(* IEC 61131-3 sources: daoli-st-library/DL_Process (part 25) *)

(* ---- FB_DL_CathodeKilnZoneSeq.st ---- *)
(*
  Component : FB_DL_CathodeKilnZoneSeq
  Category  : DL_Process
  Function  : 辊道窑多温区升温曲线执行状态机：预热→升温→保温→冷却→出料
  Complexity: C4
  开源溯源 : DLF 内部原创（R94 族模板派生）；参考语义来源见 SOURCE_HUNTING_MATRIX.md
  规则遵从 : R1-R16
  契约     : 输入 xStart 启动（上升沿启动，下降沿兼故障复位沿）、xStop 停止、xRollerOk 辊道运行正常、
             xRodBroken 断棒检测、xDischDone 出料完成、afZoneTempC 八温区实测温度定长数组 [℃]
             （ARRAY[0..7]，未用槽填零，R15 显式定长）、nZoneCount 有效温区数 [区]、
             rStartC 起始炉温 [℃]、rPreheatC 预热终点 [℃]、rSoakSetC 保温设定 [℃]、
             rRampRateKmin 升降温速率上限 [K/min]、rTempTolK 区温偏差允许带 [K]、
             rOverTempK 超温判据余量 [K]、rCoolTargetC 冷却终点 [℃]、rSoakTimeS 保温时间 [s]、
             rHeatMaxS 升温允许最长 [s]、rCoolMaxS 冷却允许最长 [s]、rDischTmoS 出料超时 [s]。
  输出     : 三路独立命令、ePhase 当前相、xFault/nFaultCode 故障、nWarnCode 信息级码、
             rZoneDevMaxK 各区相对保温设定的最大偏差 [K]、rMaxTempC/rMinTempC 区温极值 [℃]、
             xOverTemp 超温标志、xRateViol 速率越限标志。
  时序     : 同拍双窗配比约束 rHeatMaxS ≥ (rSoakSetC − rStartC) / rRampRateKmin × 60（否则升温窗
             先于工艺升温完成即超时）、rCoolMaxS ≥ (rSoakSetC − rCoolTargetC) / rRampRateKmin × 60。
  速率限幅 : 升温相以进相时刻的炉温为基准，允许温度 = 基准 + 速率 × 已用时间，实测超越即本拍断加热；
             降温相以进相时刻的炉温为基准，允许温度 = 基准 − 速率 × 已用时间，实测低于即本拍断风机。
  安全侧   : 断棒（xRodBroken）与辊道停转（NOT xRollerOk）在非待机相立即迁 FAULT 并撤销全部命令；
             断棒/停转在待机相不锁存，但阻断启动（启动条件已含两者）。
  复位沿   : 故障码锁存至 xStart 下降沿；复位后停在 IDLE，需重新给出启动上升沿才继续（不做自动再入）。
  码位     : 9820 升温速率超限（信息级）；9821 降温速率超限（信息级）；9822 区温偏差超带（信息级）；
             9823 超温转冷却（信息级）；9824 断棒（故障级）；9825 辊道停转（故障级）；
             9826 参数或温度数组非法（故障级）；9827 升温超时（故障级）；9828 冷却超时（故障级）；
             9829 出料超时（故障级）。信息级码一律不置 xFault。
*)
TYPE E_DL_KilnPhase :
(
    IDLE      := 0,    // 待机，全部命令撤销 EN: idle, every command withdrawn
    PREHEAT   := 10,   // 预热段升温 EN: the preheat ramp phase
    RAMP      := 20,   // 升温段至保温设定 EN: the ramp phase towards the soak setpoint
    SOAK      := 30,   // 保温段 EN: the soak phase
    COOL      := 40,   // 冷却段 EN: the cooling phase
    DISCHARGE := 50,   // 出料段 EN: the discharge phase
    FAULT     := 90    // 故障相，全部命令强制撤销 EN: fault phase, every command forced off
);
END_TYPE

FUNCTION_BLOCK FB_DL_CathodeKilnZoneSeq
VAR_INPUT
    xStart       : BOOL;                        // 启动（上升沿启动，下降沿复位故障） EN: start on the rising edge, reset the fault on the falling edge
    xStop        : BOOL;                        // 停止（任意相生效） EN: stop, effective in every phase
    xRollerOk    : BOOL;                        // 辊道运行正常（变频器运行反馈） EN: the roller table runs normally
    xRodBroken   : BOOL;                        // 断棒检测（安全侧信号） EN: the broken rod detection, a safety side signal
    xDischDone   : BOOL;                        // 出料完成（下游确认） EN: the discharge is complete, confirmed downstream
    afZoneTempC  : ARRAY[0..7] OF REAL;         // 八温区实测温度，未用槽填零 [℃] EN: the measured temperatures of eight zones, unused slots hold zero
    nZoneCount   : INT := 8;                    // 有效温区数 [区] EN: the number of valid zones
    rStartC      : REAL := 25.0;                // 起始炉温（升温速率基准的缺省值） [℃] EN: the starting furnace temperature used as the default ramp base
    rPreheatC    : REAL := 400.0;               // 预热终点温度 [℃] EN: the preheat end temperature
    rSoakSetC    : REAL := 800.0;               // 保温设定温度 [℃] EN: the soak setpoint temperature
    rRampRateKmin: REAL := 3.0;                 // 升降温速率上限 [K/min] EN: the upper bound of the heating and cooling rate
    rTempTolK    : REAL := 15.0;                // 区温偏差允许带 [K] EN: the allowed zone temperature deviation band
    rOverTempK   : REAL := 20.0;                // 超温判据余量（超过设定即转冷却） [K] EN: the over temperature margin above the setpoint
    rCoolTargetC : REAL := 80.0;                // 冷却终点温度 [℃] EN: the cooling end temperature
    rSoakTimeS   : REAL := 3600.0;              // 保温时间设定 [s] EN: the soak time setting
    rHeatMaxS    : REAL := 7200.0;              // 升温允许最长（预热+升温合计） [s] EN: the longest heating time covering preheat and ramp
    rCoolMaxS    : REAL := 7200.0;              // 冷却允许最长 [s] EN: the longest cooling time
    rDischTmoS   : REAL := 1800.0;              // 出料超时设定 [s] EN: the discharge timeout setting
END_VAR
VAR_OUTPUT
    xHeatCmd    : BOOL;               // 加热使能命令 EN: the heating enable command
    xFanCoolCmd : BOOL;               // 冷却风机命令 EN: the cooling fan command
    xDischCmd   : BOOL;               // 出料辊道命令 EN: the discharge conveyor command
    ePhase      : E_DL_KilnPhase;     // 当前相 EN: the current phase
    xFault      : BOOL;               // 故障标志（仅故障级码置位） EN: the fault flag, raised by fault class codes only
    nFaultCode  : INT;                // 故障码，锁存回放 EN: the fault code replayed from the latch
    nWarnCode   : INT;                // 信息级码（每拍重算） EN: the information class code recomputed every cycle
    rZoneDevMaxK: REAL;               // 各区相对保温设定的最大偏差 [K] EN: the largest zone deviation from the soak setpoint
    rMaxTempC   : REAL;               // 区温最大值 [℃] EN: the highest zone temperature
    rMinTempC   : REAL;               // 区温最小值 [℃] EN: the lowest zone temperature
    xOverTemp   : BOOL;               // 超温标志 EN: the over temperature flag
    xRateViol   : BOOL;               // 速率越限标志 EN: the rate violation flag
END_VAR
VAR
    tonHeat    : TON;                 // 升温（预热+升温）总时长定时器 EN: the total heating timer
    tonSoak    : TON;                 // 保温定时器 EN: the soak timer
    tonCool    : TON;                 // 冷却时长定时器 EN: the cooling timer
    tonDisch   : TON;                 // 出料超时定时器 EN: the discharge timeout
    fbStartRise: R_TRIG;              // xStart 上升沿（唯一启动沿） EN: the rising edge of xStart, the only start edge
    fbStartFall: F_TRIG;              // xStart 下降沿（复位沿） EN: the falling edge of xStart, the reset edge
    xFinAll    : BOOL;                // 标量浮点入参有限 EN: the scalar floating inputs are finite
    xZoneFin   : BOOL;                // 全部有效温区读数有限 EN: every valid zone reading is finite
    xParamBad  : BOOL;                // 参数或数组非法 EN: a parameter or the array is illegal
    xZoneDevOk : BOOL;                // 区温偏差在允许带内 EN: the zone deviation is inside the band
    i          : INT;                 // 温区循环索引 [区] EN: the zone loop index
    nScan      : INT;                 // 实际扫描温区数 [区] EN: the effective zone scan count
    rMax       : REAL;                // 区温最大值累加器 [℃] EN: the zone maximum accumulator
    rMin       : REAL;                // 区温最小值累加器 [℃] EN: the zone minimum accumulator
    rDev       : REAL;                // 偏差累加器 [K] EN: the deviation accumulator
    rDevMax    : REAL;                // 最大偏差 [K] EN: the largest deviation
    rHeatBaseC : REAL;                // 升温相进相基准炉温 [℃] EN: the furnace temperature latched when heating starts
    rCoolBaseC : REAL;                // 冷却相进相基准炉温 [℃] EN: the furnace temperature latched when cooling starts
    rAllowC    : REAL;                // 本拍允许温度（速率限幅） [℃] EN: the temperature allowed in this cycle by the rate limit
    rElapsedS  : REAL;                // 相内已用时间 [s] EN: the elapsed time inside the phase
    nMsSoak    : UDINT := 3600000;    // 保温毫秒数（缺省防零 PT） EN: the soak milliseconds, the default avoids a zero preset
    nMsHeat    : UDINT := 7200000;    // 升温毫秒数 EN: the heating milliseconds
    nMsCool    : UDINT := 7200000;    // 冷却毫秒数 EN: the cooling milliseconds
    nMsDisch   : UDINT := 1800000;    // 出料毫秒数 EN: the discharge milliseconds
    nCodeLatch : INT;                 // 故障码锁存副本 EN: the latched copy of the fault code
END_VAR
VAR CONSTANT
    DL_CKZ_Z      : REAL := 0.0;      // 浮点零常量 EN: the floating point zero constant
    DL_CKZ_SECMIN : REAL := 60.0;     // 分钟换算秒系数 EN: the minute to second factor
    DL_CKZ_K1000  : REAL := 1000.0;   // 秒转毫秒系数 EN: the second to millisecond factor
    DL_CKZ_IDX_MAX: INT := 7;         // 温区数组上界索引 [区] EN: the zone array upper bound index
    DL_CKZ_CNT_MAX: INT := 8;         // 温区个数上限 [区] EN: the zone count upper bound
    DL_CKZ_W_RATE : INT := 9820;      // 升温速率超限（信息级） EN: the heating rate violation, information class
    DL_CKZ_W_COOL : INT := 9821;      // 降温速率超限（信息级） EN: the cooling rate violation, information class
    DL_CKZ_W_DEV  : INT := 9822;      // 区温偏差超带（信息级） EN: the zone deviation violation, information class
    DL_CKZ_W_OVER : INT := 9823;      // 超温转冷却（信息级） EN: the over temperature transfer, information class
    DL_CKZ_C_ROD  : INT := 9824;      // 断棒（故障级） EN: the broken rod
    DL_CKZ_C_ROLL : INT := 9825;      // 辊道停转（故障级） EN: the roller table stopped
    DL_CKZ_C_PARAM: INT := 9826;      // 参数或温度数组非法（故障级） EN: a parameter or the temperature array is illegal
    DL_CKZ_C_HEAT : INT := 9827;      // 升温超时（故障级） EN: the heating timed out
    DL_CKZ_C_COOL : INT := 9828;      // 冷却超时（故障级） EN: the cooling timed out
    DL_CKZ_C_DISCH: INT := 9829;      // 出料超时（故障级） EN: the discharge timed out
END_VAR

// 段1｜参数与采样门禁：标量浮点闸 + 温区数组逐个闸（先判后用，换算在闸后）
xFinAll := (rStartC = rStartC) AND ((rStartC - rStartC) = DL_CKZ_Z)
        AND (rPreheatC = rPreheatC) AND ((rPreheatC - rPreheatC) = DL_CKZ_Z)
        AND (rSoakSetC = rSoakSetC) AND ((rSoakSetC - rSoakSetC) = DL_CKZ_Z)
        AND (rRampRateKmin = rRampRateKmin) AND ((rRampRateKmin - rRampRateKmin) = DL_CKZ_Z)
        AND (rTempTolK = rTempTolK) AND ((rTempTolK - rTempTolK) = DL_CKZ_Z)
        AND (rOverTempK = rOverTempK) AND ((rOverTempK - rOverTempK) = DL_CKZ_Z)
        AND (rCoolTargetC = rCoolTargetC) AND ((rCoolTargetC - rCoolTargetC) = DL_CKZ_Z)
        AND (rSoakTimeS = rSoakTimeS) AND ((rSoakTimeS - rSoakTimeS) = DL_CKZ_Z)
        AND (rHeatMaxS = rHeatMaxS) AND ((rHeatMaxS - rHeatMaxS) = DL_CKZ_Z)
        AND (rCoolMaxS = rCoolMaxS) AND ((rCoolMaxS - rCoolMaxS) = DL_CKZ_Z)
        AND (rDischTmoS = rDischTmoS) AND ((rDischTmoS - rDischTmoS) = DL_CKZ_Z);                        // 十一个标量入参有限性 EN: the finiteness of all eleven scalar inputs
xParamBad := (NOT xFinAll) OR (nZoneCount < 1) OR (nZoneCount > DL_CKZ_CNT_MAX)
          OR (rRampRateKmin <= DL_CKZ_Z) OR (rSoakTimeS <= DL_CKZ_Z) OR (rHeatMaxS <= DL_CKZ_Z)
          OR (rCoolMaxS <= DL_CKZ_Z) OR (rDischTmoS <= DL_CKZ_Z) OR (rTempTolK <= DL_CKZ_Z)
          OR (rOverTempK < DL_CKZ_Z) OR (rSoakSetC <= rPreheatC) OR (rPreheatC <= rStartC)
          OR (rCoolTargetC >= rSoakSetC);                                                                 // 域闸与曲线单调性约束 EN: the domain gate and the profile monotonicity
nScan := nZoneCount;                                                                                      // 扫描个数 [区] EN: the scan count
rMax := DL_CKZ_Z;                                                                                         // 最大值初值 [℃] EN: the maximum accumulator initial value
rMin := DL_CKZ_Z;                                                                                         // 最小值初值 [℃] EN: the minimum accumulator initial value
rDevMax := DL_CKZ_Z;                                                                                      // 最大偏差初值 [K] EN: the largest deviation initial value
xZoneFin := TRUE;                                                                                         // 假定温区有限 EN: assume the zones are finite
IF (nScan >= 1) AND (nScan <= DL_CKZ_CNT_MAX) THEN                                                       // 个数合法才访问数组 EN: access the array only with a legal count
    FOR i := 0 TO nScan - 1 DO                                                                           // 定长数组循环（上界已证 ≤7） EN: the fixed array loop, the bound is proven at most seven
        IF (i >= 0) AND (i <= DL_CKZ_IDX_MAX) THEN                                                       // 逐元素双边界校验 EN: the per element bound check
            IF (afZoneTempC[i] = afZoneTempC[i]) AND ((afZoneTempC[i] - afZoneTempC[i]) = DL_CKZ_Z) THEN
                IF (i = 0) OR (afZoneTempC[i] > rMax) THEN                                               // 首元素或更大值 EN: the first element or a larger value
                    rMax := afZoneTempC[i];                                                              // 更新最大值 [℃] EN: update the maximum
                END_IF
                IF (i = 0) OR (afZoneTempC[i] < rMin) THEN                                               // 首元素或更小值 EN: the first element or a smaller value
                    rMin := afZoneTempC[i];                                                              // 更新最小值 [℃] EN: update the minimum
                END_IF
                rDev := ABS(afZoneTempC[i] - rSoakSetC);                                                 // 相对保温设定的偏差 [K] EN: the deviation from the soak setpoint
                IF rDev > rDevMax THEN                                                                   // 取更大偏差 EN: keep the larger deviation
                    rDevMax := rDev;                                                                     // 更新最大偏差 [K] EN: update the largest deviation
                END_IF
            ELSE
                xZoneFin := FALSE;                                                                       // 记非有限元素 EN: mark the non finite element
            END_IF
        END_IF
    END_FOR
ELSE
    xZoneFin := FALSE;                                                                                   // 个数非法等同读数不可用 EN: an illegal count makes the readings unusable
END_IF
xParamBad := xParamBad OR (NOT xZoneFin);                                                                // 读数不可用并入参数闸（单点写入） EN: merge the unusable readings into the parameter gate
IF (NOT xParamBad) THEN                                                                                  // 参数合法才做时间换算 EN: convert only when the parameters are legal
    nMsSoak := REAL_TO_UDINT(rSoakTimeS * DL_CKZ_K1000);                                                 // 保温毫秒数 EN: the soak milliseconds
    nMsHeat := REAL_TO_UDINT(rHeatMaxS * DL_CKZ_K1000);                                                  // 升温毫秒数 EN: the heating milliseconds
    nMsCool := REAL_TO_UDINT(rCoolMaxS * DL_CKZ_K1000);                                                  // 冷却毫秒数 EN: the cooling milliseconds
    nMsDisch := REAL_TO_UDINT(rDischTmoS * DL_CKZ_K1000);                                                // 出料毫秒数 EN: the discharge milliseconds
END_IF
xZoneDevOk := (NOT xParamBad) AND (rDevMax <= rTempTolK);                                                // 区温偏差带内判据 EN: the zone deviation band test

// 段2｜四只定时器 + 两只边沿实例无条件周期刷新（CASE 内不调用实例）
tonHeat(IN := (ePhase = E_DL_KilnPhase.PREHEAT) OR (ePhase = E_DL_KilnPhase.RAMP), PT := UDINT_TO_TIME(nMsHeat));  // 升温总时长 EN: the total heating time
tonSoak(IN := (ePhase = E_DL_KilnPhase.SOAK) AND xZoneDevOk, PT := UDINT_TO_TIME(nMsSoak));                          // 保温计时（偏差在带内才累计） EN: count the soak only inside the band
tonCool(IN := (ePhase = E_DL_KilnPhase.COOL), PT := UDINT_TO_TIME(nMsCool));                                         // 冷却时长 EN: the cooling time
tonDisch(IN := (ePhase = E_DL_KilnPhase.DISCHARGE), PT := UDINT_TO_TIME(nMsDisch));                                  // 出料时长 EN: the discharge time
fbStartRise(CLK := xStart);                                                                                          // 启动沿 EN: the start edge
fbStartFall(CLK := xStart);                                                                                          // 复位沿 EN: the reset edge

// 段3｜输出预置（唯一预置点，CASE 内只置位；信息级码每拍重算）
xHeatCmd := FALSE;                        // 加热预置关 EN: preset the heating off
xFanCoolCmd := FALSE;                     // 风机预置停 EN: preset the fan off
xDischCmd := FALSE;                       // 出料预置停 EN: preset the discharge off
xFault := FALSE;                          // 故障标志预置假 EN: preset the fault flag false
nFaultCode := 0;                          // 故障码预置零 EN: preset the fault code to zero
nWarnCode := 0;                           // 信息码预置零 EN: preset the warning code to zero
xOverTemp := FALSE;                       // 超温标志预置假 EN: preset the over temperature flag false
xRateViol := FALSE;                       // 速率越限标志预置假 EN: preset the rate violation flag false
rZoneDevMaxK := rDevMax;                  // 最大偏差出口 [K] EN: publish the largest deviation
rMaxTempC := rMax;                        // 区温最大值出口 [℃] EN: publish the highest zone temperature
rMinTempC := rMin;                        // 区温最小值出口 [℃] EN: publish the lowest zone temperature

// 段4｜全局安全闸：参数非法 / 断棒 / 辊道停转 → 锁故障；xStop 撤销命令回待机
IF xParamBad THEN
    nCodeLatch := DL_CKZ_C_PARAM;                                                                        // 参数非法锁存 EN: latch the parameter code
    xFault := TRUE;                                                                                      // 置故障标志 EN: raise the fault flag
    nFaultCode := DL_CKZ_C_PARAM;                                                                        // 故障码出口 EN: publish the fault code
    ePhase := E_DL_KilnPhase.FAULT;                                                                      // 迁故障相 EN: move to the fault phase
ELSIF xRodBroken AND (ePhase <> E_DL_KilnPhase.IDLE) THEN
    nCodeLatch := DL_CKZ_C_ROD;                                                                          // 断棒锁存 EN: latch the broken rod code
    xFault := TRUE;                                                                                      // 置故障标志 EN: raise the fault flag
    nFaultCode := DL_CKZ_C_ROD;                                                                          // 故障码出口 EN: publish the fault code
    ePhase := E_DL_KilnPhase.FAULT;                                                                      // 迁故障相 EN: move to the fault phase
ELSIF (NOT xRollerOk) AND (ePhase <> E_DL_KilnPhase.IDLE) THEN
    nCodeLatch := DL_CKZ_C_ROLL;                                                                         // 辊道停转锁存 EN: latch the roller stop code
    xFault := TRUE;                                                                                      // 置故障标志 EN: raise the fault flag
    nFaultCode := DL_CKZ_C_ROLL;                                                                         // 故障码出口 EN: publish the fault code
    ePhase := E_DL_KilnPhase.FAULT;                                                                      // 迁故障相 EN: move to the fault phase
ELSIF xStop AND (ePhase <> E_DL_KilnPhase.IDLE) THEN
    ePhase := E_DL_KilnPhase.IDLE;                                                                       // 撤销型停车回待机 EN: a withdrawing stop returns to idle
END_IF

// 段5｜主状态机（ENUM + CASE，ELSE 兜底非法值）
IF ePhase <> E_DL_KilnPhase.FAULT THEN
CASE ePhase OF
E_DL_KilnPhase.IDLE:
    // 拍 N：待机；启动需辊道正常、无断棒、无停车（入相即锁存速率限幅基准炉温）
    IF fbStartRise.Q AND xRollerOk AND (NOT xRodBroken) AND (NOT xStop) AND (NOT xParamBad) THEN
        rHeatBaseC := rMax;                                                                              // 锁存升温基准炉温 [℃] EN: latch the heating base temperature
        ePhase := E_DL_KilnPhase.PREHEAT;                                                                // 本拍行为：进预热相 EN: enter the preheat phase
    END_IF

E_DL_KilnPhase.PREHEAT:
    // 拍 N：预热升温，速率越限即本拍断加热（信息级 9820），升到预热终点转升温相
    rElapsedS := TIME_TO_REAL(tonHeat.ET) * 0.001;                                                       // 已用时间 [s] EN: the elapsed time
    rAllowC := rHeatBaseC + rRampRateKmin * (rElapsedS / DL_CKZ_SECMIN);                                 // 允许温度 [℃] EN: the temperature allowed by the rate limit
    IF rMax > (rAllowC + rTempTolK) THEN                                                                 // 速率越限判据 EN: the rate violation test
        xRateViol := TRUE;                                                                               // 置越限标志 EN: raise the rate flag
        nWarnCode := DL_CKZ_W_RATE;                                                                      // 信息级码，不置故障 EN: an information class code, no fault
    ELSE
        xHeatCmd := TRUE;                                                                                // 加热允许 EN: heating allowed
    END_IF
    IF rMax >= rPreheatC THEN                                                                            // 预热到位 EN: the preheat is complete
        ePhase := E_DL_KilnPhase.RAMP;                                                                   // 本拍行为：进升温相 EN: enter the ramp phase
    ELSIF tonHeat.Q THEN
        nCodeLatch := DL_CKZ_C_HEAT;                                                                     // 升温超时 EN: the heating timed out
        xFault := TRUE;                                                                                  // 置故障标志 EN: raise the fault flag
        nFaultCode := DL_CKZ_C_HEAT;                                                                     // 故障码出口 EN: publish the fault code
        ePhase := E_DL_KilnPhase.FAULT;                                                                  // 迁故障相 EN: move to the fault phase
    END_IF

E_DL_KilnPhase.RAMP:
    // 拍 N：升温至保温设定，含速率限幅与升温超时兜底
    rElapsedS := TIME_TO_REAL(tonHeat.ET) * 0.001;                                                       // 已用时间（含预热相） [s] EN: the elapsed time including the preheat phase
    rAllowC := rHeatBaseC + rRampRateKmin * (rElapsedS / DL_CKZ_SECMIN);                                 // 允许温度 [℃] EN: the allowed temperature
    IF rMax > (rAllowC + rTempTolK) THEN                                                                 // 速率越限判据 EN: the rate violation test
        xRateViol := TRUE;                                                                               // 置越限标志 EN: raise the rate flag
        nWarnCode := DL_CKZ_W_RATE;                                                                      // 信息级码 EN: the information class code
    ELSE
        xHeatCmd := TRUE;                                                                                // 加热允许 EN: heating allowed
    END_IF
    IF rMax >= (rSoakSetC - rTempTolK) THEN                                                              // 到达保温窗口下沿 EN: reached the lower edge of the soak window
        ePhase := E_DL_KilnPhase.SOAK;                                                                   // 本拍行为：进保温相 EN: enter the soak phase
    ELSIF tonHeat.Q THEN
        nCodeLatch := DL_CKZ_C_HEAT;                                                                     // 升温超时 EN: the heating timed out
        xFault := TRUE;                                                                                  // 置故障标志 EN: raise the fault flag
        nFaultCode := DL_CKZ_C_HEAT;                                                                     // 故障码出口 EN: publish the fault code
        ePhase := E_DL_KilnPhase.FAULT;                                                                  // 迁故障相 EN: move to the fault phase
    END_IF

E_DL_KilnPhase.SOAK:
    // 拍 N：保温；超温立即转冷却（信息级 9823），偏差超带只告警（9822）且不累计保温时间
    IF rMax > (rSoakSetC + rOverTempK) THEN                                                              // 超温判据 EN: the over temperature test
        xOverTemp := TRUE;                                                                               // 置超温标志 EN: raise the over temperature flag
        nWarnCode := DL_CKZ_W_OVER;                                                                      // 超温信息级码 EN: the over temperature information code
        rCoolBaseC := rMin;                                                                              // 锁存冷却基准炉温 [℃] EN: latch the cooling base temperature
        ePhase := E_DL_KilnPhase.COOL;                                                                   // 本拍行为：立即转冷却 EN: transfer to cooling immediately
    ELSIF NOT xZoneDevOk THEN
        nWarnCode := DL_CKZ_W_DEV;                                                                       // 偏差超带告警（信息级） EN: warn about the zone deviation
        xHeatCmd := TRUE;                                                                                // 保持加热以拉回设定 EN: keep heating to recover the setpoint
    ELSE
        xHeatCmd := TRUE;                                                                                // 保温加热 EN: soak heating
        IF tonSoak.Q THEN                                                                                // 保温时间到 EN: the soak time elapsed
            rCoolBaseC := rMin;                                                                          // 锁存冷却基准炉温 [℃] EN: latch the cooling base temperature
            ePhase := E_DL_KilnPhase.COOL;                                                               // 本拍行为：进冷却相 EN: enter the cooling phase
        END_IF
    END_IF

E_DL_KilnPhase.COOL:
    // 拍 N：冷却；降温过快本拍断风机（信息级 9821），降到终点转出料，冷却超时判 9828
    rElapsedS := TIME_TO_REAL(tonCool.ET) * 0.001;                                                       // 冷却已用时间 [s] EN: the cooling elapsed time
    rAllowC := rCoolBaseC - rRampRateKmin * (rElapsedS / DL_CKZ_SECMIN);                                 // 允许温度（速率下限） [℃] EN: the allowed temperature floor
    IF rMin < (rAllowC - rTempTolK) THEN                                                                 // 降温超速率判据 EN: the over fast cooling test
        xRateViol := TRUE;                                                                               // 置越限标志 EN: raise the rate flag
        nWarnCode := DL_CKZ_W_COOL;                                                                      // 信息级码 EN: the information class code
    ELSE
        xFanCoolCmd := TRUE;                                                                             // 风机允许 EN: the fan is allowed
    END_IF
    IF rMax <= rCoolTargetC THEN                                                                         // 冷却到位 EN: the cooling is complete
        ePhase := E_DL_KilnPhase.DISCHARGE;                                                              // 本拍行为：进出料相 EN: enter the discharge phase
    ELSIF tonCool.Q THEN
        nCodeLatch := DL_CKZ_C_COOL;                                                                     // 冷却超时 EN: the cooling timed out
        xFault := TRUE;                                                                                  // 置故障标志 EN: raise the fault flag
        nFaultCode := DL_CKZ_C_COOL;                                                                     // 故障码出口 EN: publish the fault code
        ePhase := E_DL_KilnPhase.FAULT;                                                                  // 迁故障相 EN: move to the fault phase
    END_IF

E_DL_KilnPhase.DISCHARGE:
    // 拍 N：出料；下游确认回待机，超时判 9829（迁入本相已带参数闸复检）
    IF xDischDone THEN                                                                                   // 出料完成 EN: the discharge is complete
        ePhase := E_DL_KilnPhase.IDLE;                                                                   // 本拍行为：回待机 EN: back to idle
    ELSIF tonDisch.Q THEN
        nCodeLatch := DL_CKZ_C_DISCH;                                                                    // 出料超时 EN: the discharge timed out
        xFault := TRUE;                                                                                  // 置故障标志 EN: raise the fault flag
        nFaultCode := DL_CKZ_C_DISCH;                                                                    // 故障码出口 EN: publish the fault code
        ePhase := E_DL_KilnPhase.FAULT;                                                                  // 迁故障相 EN: move to the fault phase
    END_IF

E_DL_KilnPhase.FAULT:
    // 故障相（本段被外层 IF 排除，保留分支以满足枚举穷举）
    xFault := TRUE;                                                                                      // 保持故障标志 EN: keep the fault flag
    nFaultCode := nCodeLatch;                                                                            // 锁存回放 EN: replay the latch

ELSE
    // 非法状态兜底：绝不停在未知相
    nCodeLatch := DL_CKZ_C_PARAM;                                                                        // 非法状态归参数码 EN: treat an illegal state as a parameter code
    xFault := TRUE;                                                                                      // 置故障标志 EN: raise the fault flag
    nFaultCode := DL_CKZ_C_PARAM;                                                                        // 故障码出口 EN: publish the fault code
    ePhase := E_DL_KilnPhase.FAULT;                                                                      // 迁故障相 EN: move to the fault phase
END_CASE
END_IF

// 段6｜相独立使能出口（IDLE/FAULT 不置任何命令，天然强制撤销；出料相另给辊道命令）
CASE ePhase OF
E_DL_KilnPhase.DISCHARGE:
    xDischCmd := TRUE;                                                                                   // 出料辊道命令 EN: the discharge conveyor command
ELSE
    xDischCmd := FALSE;                                                                                  // 其余相撤销出料命令 EN: withdraw the discharge command elsewhere
END_CASE

// 段7｜故障相锁存回放 + 复位沿（xStart 下降沿清除，复位后停 IDLE 需重新给启动上升沿）
IF ePhase = E_DL_KilnPhase.FAULT THEN
    xFault := TRUE;                                                                                      // 故障标志保持 EN: keep the fault flag
    nFaultCode := nCodeLatch;                                                                            // 锁存回放，不按当下输入重推断 EN: replay the latch instead of re inferring
    nWarnCode := 0;                                                                                      // 故障相不报信息级码 EN: no information class code in the fault phase
    xHeatCmd := FALSE;                                                                                   // 加热强制关 EN: force the heating off
    xFanCoolCmd := FALSE;                                                                                // 风机强制停（断棒时避免热冲击） EN: force the fan off to avoid a thermal shock
    xDischCmd := FALSE;                                                                                  // 出料强制停 EN: force the discharge off
    IF fbStartFall.Q THEN
        nCodeLatch := 0;                                                                                 // 清除边：xStart 下降沿（头注释已声明） EN: clear on the falling edge of xStart
        ePhase := E_DL_KilnPhase.IDLE;                                                                   // 回待机 EN: back to idle
    END_IF
END_IF
END_FUNCTION_BLOCK

(* ---- FB_DL_CellAgingRestSeq.st ---- *)
(*
  组件名 Component   : FB_DL_CellAgingRestSeq
  子库 Sublibrary    : DL_Process
  版本 Version       : 1.0.0
  兼容性 Platform    : CODESYS 3.5 / TwinCAT 3 / 汇川 InoProShop / Machine Expert（仅 Standard.library）
  功能 Function      : 电芯老化静置顺控（自研行业池：锂电）：
                       1) 静置计时：tRestDur 总静置时长承载（独立 TON）；
                       2) 抽测窗口：静置相内周期开抽测窗（周期计 tonSampleInt 自复触，
                       R188），窗长 tSampleWin；窗口结束后锁存最后一次抽测值；
                       3) 时限到期判级出柜：静置时长到 → 按末次抽测电压与内阻判级
                       （合格 ePass / 降级 eMarginal / 不合格 eFail），结果锁存至复位；
                       4) 静置中断判据：抽测窗内电压越域持续 tVoltDevTo → 故障锁存。
  边界 Boundary      : ① 本件只出抽测请求与判级结论，不驱动充放电（老化柜本体自控）；
                       ② 判级只认末次抽测锁存值（禁按当下输入重推断，R152）；
                       ③ 周期窗计时自复触范式（R188），静置/窗口/越带确认独立实例；
                       ④ 故障锁存解除唯一路径 = bReset 上升沿（输入引脚，恒可达）；
                       ⑤ 无全局变量引用、无外部变量声明、无物理地址寻址。
  依赖 Depends       : Standard.library（R_TRIG / TON）
  溯源 Origin        : 道莅自研 clean-room（自研行业池：锂电老化静置共性语义，
                       零外部代码行复制）
  码位 Code          : 16#06_0_C0（Process 段 0006，C 子带 C0 格）
  码表 Error codes（本件格 06_0_C0，单轨子道：故障 0x02C0 / 信息 0x01C0）:
    16#0006_02C0 故障级：静置顺控故障总码（电压越域 / 组态非法 / 输入非有限），
                 锁存至复位
    16#0006_01C0 信息级：判级完成沿（ePass/eMarginal/eFail 写定拍）
  修订历史 Revision  :
    2026-11-19  v1.0.0  R44 首版（批次 4 · 序号 17）
*)

TYPE E_DL_CarPhase :
(
    eIdle     := 0,   // 空闲：未使能 / Idle, not enabled
    eRest     := 10,  // 静置：计时 + 周期抽测 / Resting with periodic sampling
    eSample   := 20,  // 抽测：窗口驻留 / Sampling window dwell
    eGrade    := 30,  // 判级：末次抽测定级 / Grading from last sample
    eDone     := 40,  // 完成：结论驻留 / Done, verdict held
    eFault    := 90   // 故障：总码锁存 / Fault, latched
);
END_TYPE

TYPE E_DL_CarGrade :
(
    eNone     := 0,   // 无结论 / No verdict
    ePass     := 10,  // 合格：电压内阻双达标 / Pass
    eMarginal := 20,  // 降级：电压入降级带 / Marginal
    eFail     := 30   // 不合格：越降级带下限或内阻不足 / Fail
);
END_TYPE

FUNCTION_BLOCK FB_DL_CellAgingRestSeq
VAR_INPUT
    bEnable     : BOOL;                  // 使能（电平）[-] / Enable
    bReset      : BOOL;                  // 上升沿清故障锁存 [-] / Reset edge
    fCellVoltV  : REAL;                  // 电芯实测电压 [伏特] / Cell voltage
    fIrMohm     : REAL;                  // 电芯实测内阻 [毫欧] / Internal resistance
    tRestDur    : TIME := T#72H;         // 总静置时长 [毫秒] / Total rest duration
    tSampleInt  : TIME := T#4H;          // 抽测周期 [毫秒] / Sample interval
    tSampleWin  : TIME := T#60S;         // 抽测窗口长 [毫秒] / Sample window duration
    fVoltPassLoV: REAL := 3.60;          // 合格电压下限 [伏特] / Pass voltage floor
    fVoltMargLoV: REAL := 3.50;          // 降级电压下限 [伏特] / Marginal voltage floor
    fIrMinMohm  : REAL := 1.0;           // 合格内阻下限 [毫欧] / IR pass floor
    tVoltDevTo  : TIME := T#10S;         // 电压越域确认窗 [毫秒] / Voltage deviation timeout
END_VAR
VAR_OUTPUT
    bSampleReq  : BOOL;                  // 抽测请求电平（窗口相）[-] / Sample request level
    fVoltLastV  : REAL;                  // 末次抽测电压 [伏特] / Last sampled voltage
    fIrLastMohm : REAL;                  // 末次抽测内阻 [毫欧] / Last sampled IR
    eGrade      : E_DL_CarGrade;         // 判级结论出口 / Grade verdict outlet
    ePhase      : E_DL_CarPhase;         // 相位出口，段尾单点映射 / Phase outlet
    bError      : BOOL;                  // 故障锁存标志 [-] / Fault latch flag
    uErrId      : UDINT;                 // 事件码，0 = 无事件 / Event code
END_VAR
VAR
    rtReset    : R_TRIG;                 // 复位沿实例，段 0 无条件刷新 / Reset edge
    tonRestDur : TON;                    // 静置总时长计时（独立实例） / Rest duration timer
    tonSampleInt: TON;                   // 抽测周期计（自复触，R188） / Sample interval timer
    tonSampleWin: TON;                   // 抽测窗口计时（独立实例） / Sample window timer
    tonVoltDevTo: TON;                   // 电压越域确认（专用超时件命名） / Voltage timeout
    _ePhase    : E_DL_CarPhase := E_DL_CarPhase.eIdle;    // 内部相位（CASE 唯一写入目标）/ Internal phase
    _eGrade    : E_DL_CarGrade := E_DL_CarGrade.eNone;    // 内部判级（锁存量）/ Internal grade
    _bFault    : BOOL;                   // 故障锁存位（锁存量） / Latched fault bit
    _uFault    : UDINT;                  // 故障码锁存（锁存量） / Latched fault code
    _bCfgBad   : BOOL;                   // 组态非法当拍量 [-] / Config illegal flag
    _bNonFin   : BOOL;                   // 输入非有限当拍量 [-] / Non-finite input flag
END_VAR
VAR CONSTANT
    DL_ABS_MAX : REAL := 1.0E30;         // 有限值判定上界 [工程单位] / Finite bound
    DL_ZERO    : REAL := 0.0;            // 零常量 [工程单位] / Zero constant
END_VAR

(* —— 段 0｜沿与定时器每拍无条件刷新（禁置于 IF/CASE 内；各实例独立禁复用） —— *)
rtReset(CLK := bReset);
tonRestDur (IN := (_ePhase = E_DL_CarPhase.eRest) AND (NOT _bFault), PT := tRestDur);
tonSampleInt(IN := (_ePhase = E_DL_CarPhase.eRest) AND (NOT _bFault) AND (NOT tonSampleInt.Q),
             PT := tSampleInt);          // 自复触周期窗：Q 拍断开一拍（R188）
tonSampleWin(IN := (_ePhase = E_DL_CarPhase.eSample) AND (NOT _bFault), PT := tSampleWin);
tonVoltDevTo(IN := (_ePhase = E_DL_CarPhase.eSample) AND ((fCellVoltV > fVoltPassLoV)
              OR (fCellVoltV < fVoltMargLoV)) AND (NOT _bFault), PT := tVoltDevTo);

(* —— 段 1｜瞬时量预清零（锁存量 _bFault/_uFault/_eGrade/fVoltLastV/fIrLastMohm 不入清单） —— *)
uErrId   := 16#0000_0000;
bSampleReq := FALSE;
_bCfgBad := FALSE;
_bNonFin := FALSE;

(* —— 段 2｜复位沿：故障与判级一次性清干净，相位回空闲 —— *)
IF rtReset.Q THEN
    _bFault := FALSE;
    _uFault := 16#0000_0000;
    _eGrade := E_DL_CarGrade.eNone;
    _ePhase := E_DL_CarPhase.eIdle;
END_IF

(* —— 段 3｜组态闸与非有限判据（覆盖全部参与判据换算引脚） —— *)
IF (fVoltMargLoV >= fVoltPassLoV) OR (fIrMinMohm <= DL_ZERO) OR (tRestDur = T#0S)
   OR (tSampleInt = T#0S) OR (tSampleWin = T#0S) OR (tVoltDevTo = T#0S) THEN
    _bCfgBad := TRUE;
END_IF
IF (fCellVoltV <> fCellVoltV) OR ((fCellVoltV - fCellVoltV) <> DL_ZERO)
   OR (fIrMohm <> fIrMohm) OR ((fIrMohm - fIrMohm) <> DL_ZERO) THEN
    _bNonFin := TRUE;
END_IF

(* —— 段 4｜主状态机：六态全覆盖 + ELSE 兜底 —— *)
CASE _ePhase OF

E_DL_CarPhase.eIdle:
    IF bEnable AND (NOT _bCfgBad) THEN
        _ePhase := E_DL_CarPhase.eRest;
    ELSIF bEnable AND _bCfgBad THEN
        _bFault := TRUE;
        _uFault := 16#0006_02C0;
        bError  := TRUE;
        _ePhase := E_DL_CarPhase.eFault;
    END_IF

E_DL_CarPhase.eRest:
    IF _bNonFin THEN
        _bFault := TRUE;
        _uFault := 16#0006_02C0;
        bError  := TRUE;
        _ePhase := E_DL_CarPhase.eFault;
    ELSIF NOT bEnable THEN
        _ePhase := E_DL_CarPhase.eIdle;  // 使能撤销回空闲
    ELSIF tonSampleInt.Q THEN
        _ePhase := E_DL_CarPhase.eSample;    // 抽测周期到：开抽测窗
    ELSIF tonRestDur.Q THEN
        _ePhase := E_DL_CarPhase.eGrade;     // 静置时长到：进判级相
    END_IF

E_DL_CarPhase.eSample:
    bSampleReq := TRUE;                  // 抽测请求电平（窗口相电平）
    IF _bNonFin THEN
        _bFault := TRUE;
        _uFault := 16#0006_02C0;
        bError  := TRUE;
        _ePhase := E_DL_CarPhase.eFault;
    ELSIF tonVoltDevTo.Q THEN
        _bFault := TRUE;                 // 窗内电压越域持续：锁存
        _uFault := 16#0006_02C0;
        bError  := TRUE;
        _ePhase := E_DL_CarPhase.eFault;
    ELSIF tonSampleWin.Q THEN
        fVoltLastV := fCellVoltV;        // 窗口结束：末次抽测值锁存（R152）
        fIrLastMohm := fIrMohm;
        bSampleReq := FALSE;
        _ePhase := E_DL_CarPhase.eRest;  // 回静置相（抽测周期重新起算）
    END_IF

E_DL_CarPhase.eGrade:
    (* 判级只认末次抽测锁存值（禁按当下输入重推断） *)
    IF (fVoltLastV >= fVoltPassLoV) AND (fIrLastMohm >= fIrMinMohm) THEN
        _eGrade := E_DL_CarGrade.ePass;  // 合格：双达标
    ELSIF (fVoltLastV >= fVoltMargLoV) AND (fIrLastMohm >= fIrMinMohm) THEN
        _eGrade := E_DL_CarGrade.eMarginal;      // 降级：电压入降级带
    ELSE
        _eGrade := E_DL_CarGrade.eFail;  // 不合格：越降级带或内阻不足
    END_IF
    uErrId := 16#0006_01C0;              // 信息级：判级完成沿
    _ePhase := E_DL_CarPhase.eDone;

E_DL_CarPhase.eDone:
    ;                                    // 结论锁存驻留（eGrade 出口回放），等复位或使能撤销
    IF NOT bEnable THEN
        _ePhase := E_DL_CarPhase.eIdle;  // 使能撤销回空闲（待机可返回路径）
    END_IF

E_DL_CarPhase.eFault:
    bError := TRUE;                      // 故障相驻留：判级与抽测值冻结，只认复位沿（段 2 迁出）
    ;                                    // （冻结语义：fVoltLastV/fIrLastMohm/_eGrade 保持）

ELSE
    _bFault := TRUE;                     // 兜底：非法相位锁存
    _uFault := 16#0006_02C0;
    bError  := TRUE;
    _ePhase := E_DL_CarPhase.eFault;
END_CASE

(* —— 段 5｜相位与判级出口单点映射（名实同源） —— *)
eGrade := _eGrade;
ePhase := _ePhase;
END_FUNCTION_BLOCK

(* ---- FB_DL_CellOcvBinSort.st ---- *)
(*
  FB_DL_CellOcvBinSort  —  OCV 分选档位落 bin（档位映射 + 满 bin 换道） / OCV bin sorting with grade mapping and full-bin lane change
  分类 Category : DL_Process
  版本 Version  : 1.0.0
  来源 Source   : roadmap-li-p1 — 锂电 OCV 分选工站真缺口
  溯源 Origin   : 道莅 clean-room 实现；四档电压阈值映射 + 落料计时 + 满 bin 换道停机为公开分选工艺逻辑，未复制任何源码行
  功能 Function : 1) 档位映射：fOcvMv 按 fTh1Mv~fTh4Mv 四阶梯阈值映射到档位 1~4
                  （阈值默认升序，第 4 档为 >= 阈值兜底档）；2) 落料相 eDispatch 由 tDrop 计时；
                  3) 档位 bin 计数 nBinUsed[档位] 递增，达 nBinCap 即 bBinFull 置位并在
                  段 3 以 03A1 锁存（满 bin 换道请求，须人工清空后复位）；
                  4) 故障级单码 03A1，归因由 eCause 独立成员承载（R190）；
                  5) 信息级 04C9 = 单件分选完成沿；6) 解除式全当拍量（R240）。
  接口 Interface: 输入 OCV 电压 + 四阈 + 容量 + 落料时间；输出状态/档位/各 bin 计数/码
  边界 Boundary : ① 组态闸：四阈值非严格升序（fTh2Mv <= fTh1Mv 等）、nBinCap = 0、
                  tDrop <= T#0S 任一成立 → 03A1 锁存；
                  ② 档位数组下标写前显式钳制（nGrade 落在 1..4，越界不写，ELSE 兜底归 4 档）；
                  ③ 浮点阈值判据为「>=」单侧直比（阈值本身无容差语义，避免误判），电压量纲
                  mV 整数化输入；④ 落料 TON 与 R_TRIG 段 0 无条件周期调用；
                  ⑤ 故障相迁出唯一路径 = bReset 上升沿；⑥ 零全局耦合（无 GVL / %I %Q %M）。
  依赖 Depends  : Standard.library（TON / R_TRIG）
  码表 Error codes（Process 段 0005，故障窗口 03A1 / 信息窗口 04C9）:
    16#0005_03A1 故障级：分选故障总码（组态非法 / 落料超时 / 目标 bin 已满需换道），
                 锁存至 bReset 上升沿；归因见 eCause，不新增码位（派单硬约束单码）
    16#0005_04C9 信息级：单件分选完成沿（落料完成计数后单拍）
  修订历史 Revision :
    2026-11-19  v1.0.0  R43 首版（批次 1 · 序号 5）
*)

TYPE E_DL_OcvState :
(
    eIdle     := 0,   // 未使能待启动 / Idle, waiting start
    eClassify := 10,  // 档位判定中 / Grade classification
    eDispatch := 20,  // 落料中（落料计时） / Dispatching with drop timer
    eDone     := 50,  // 单件完成 / Single piece done
    eFault    := 90   // 故障锁存相 / Fault latched phase
);
END_TYPE

TYPE E_DL_OcvCause :
(
    eNone       := 0, // 无故障成因 / No cause
    eCfgIllegal := 1, // 组态非法 / Illegal configuration
    eDropTmo    := 2, // 落料超时 / Drop timeout
    eBinFull    := 3  // 目标 bin 已满（换道请求） / Target bin full, lane change
);
END_TYPE

FUNCTION_BLOCK FB_DL_CellOcvBinSort
VAR_INPUT
    fOcvMv      : REAL := 0.0;        // 单体 OCV 电压 [mV] / Cell OCV voltage
    fTh1Mv      : REAL := 3300.0;     // 1/2 档分界阈值 [mV] / Grade 1-2 threshold
    fTh2Mv      : REAL := 3350.0;     // 2/3 档分界阈值 [mV] / Grade 2-3 threshold
    fTh3Mv      : REAL := 3400.0;     // 3/4 档分界阈值 [mV] / Grade 3-4 threshold
    fTh4Mv      : REAL := 3450.0;     // 4 档上界（>= 归 4 档） [mV] / Grade 4 upper threshold
    nBinCap     : UINT := 500;        // 单 bin 容量 [件]，域 > 0 / Bin capacity
    tDrop       : TIME := T#800MS;    // 落料时长 [ms]，域 > 0 / Drop duration
    bStart      : BOOL := FALSE;      // 启动命令（电平）[-] / Start command
    bBinCleared : BOOL := FALSE;      // bin 已清空确认（电平）[-] / Bin cleared acknowledge
    bReset      : BOOL := FALSE;      // 复位命令，上升沿清故障 [-] / Reset edge
END_VAR
VAR_OUTPUT
    eState      : E_DL_OcvState;      // 状态出口，段 6 单点映射 / State outlet
    eCause      : E_DL_OcvCause;      // 故障成因出口（R190） / Fault cause outlet
    nGrade      : UINT;               // 当前档位 0~4，0 = 未判定 / Current grade
    anBinUsed   : ARRAY[1..4] OF UDINT;   // 各档 bin 已用计数 [件] / Per-grade bin usage
    bBinFull    : BOOL;               // 满 bin 标志镜像 [-] / Bin full mirror
    bCycleDone  : BOOL;               // 单件完成标志 [-] / Piece done flag
    bError      : BOOL;               // 故障锁存标志 [-] / Fault latch flag
    nErrId      : UDINT;              // 事件码，0 = 无事件 / Event code
END_VAR
VAR
    _eState     : E_DL_OcvState := E_DL_OcvState.eIdle;   // 内部相位（CASE 唯一写入目标） / Internal phase
    _eCause     : E_DL_OcvCause := E_DL_OcvCause.eNone;   // 故障成因锁存（锁存量） / Latched cause
    tonDrop     : TON;                // 落料计时实例，每周期无条件调用 / Drop timer
    rtReset     : R_TRIG;             // 复位沿实例，每周期无条件调用 / Reset edge
    _anBinUsed  : ARRAY[1..4] OF UDINT;   // 内部 bin 计数（持久，段 6 映射） / Internal bin usage
    _nGrade     : UINT;               // 档位判定结果（当拍量） / Grade verdict
    _bCfgBad    : BOOL;               // 组态非法当拍量 [-] / Config illegal
    _bFault     : BOOL;               // 故障锁存位（锁存量） / Latched fault bit
    _uFault     : UDINT;              // 故障码锁存（锁存量） / Latched fault code
    _uInfo      : UDINT;              // 信息码，每拍重算 / Transient info code
END_VAR

(* —— 段 0：沿实例与定时器无条件周期刷新 + 档位判定（纯函数式，无副作用） —— *)
IF fOcvMv < fTh1Mv THEN                        // 低于 1/2 分界：1 档 / Below first threshold: grade 1
    _nGrade := 1;
ELSIF fOcvMv < fTh2Mv THEN                     // 低于 2/3 分界：2 档 / Grade 2
    _nGrade := 2;
ELSIF fOcvMv < fTh3Mv THEN                     // 低于 3/4 分界：3 档 / Grade 3
    _nGrade := 3;
ELSE                                           // 兜底：>= 3/4 分界归 4 档 / Fallback grade 4
    _nGrade := 4;
END_IF
_bCfgBad := (fTh2Mv <= fTh1Mv) OR (fTh3Mv <= fTh2Mv) OR (fTh4Mv <= fTh3Mv)
            OR (nBinCap = 0) OR (tDrop <= T#0S);                   // 组态非法当拍量 / Config illegal
rtReset(CLK := bReset);                                            // 复位沿，每拍必调 / Reset edge
tonDrop(IN := (_eState = E_DL_OcvState.eDispatch), PT := tDrop);   // 落料计时 / Drop timer

(* —— 段 1：单拍量预清零（锁存量与 bin 计数均不入清单） —— *)
_uInfo := 16#0000_0000;            // 信息码每拍重算 / Info recomputed
nGrade := 0;                       // 档位出口缺省 0 / Grade default
bBinFull := FALSE;                 // 满 bin 镜像缺省 FALSE / Bin full default
bCycleDone := FALSE;               // 完成标志缺省 FALSE / Done default
nErrId := 16#0000_0000;            // 事件码缺省无事件 / Event code default

(* —— 段 2：复位沿 + 组态域闸 —— *)
IF rtReset.Q THEN                              // rtReset.Q = 当拍量 / current scan
    _bFault := FALSE;                          // 清故障锁存位（锁存量） / Clear fault latch
    _uFault := 16#0000_0000;                   // 清故障锁存码（锁存量） / Clear fault code
    _eCause := E_DL_OcvCause.eNone;            // 清成因（锁存量） / Clear cause
    IF _eState = E_DL_OcvState.eFault THEN
        _eState := E_DL_OcvState.eIdle;        // 故障相迁出：回未使能 / Fault exit to idle
    END_IF
END_IF
IF _bCfgBad THEN                               // 组态域闸 / Config gate
    _uFault := 16#0005_03A1;                   // 故障级：分选故障总码 / Process fault code
    _eCause := E_DL_OcvCause.eCfgIllegal;      // 归因：组态非法 / Cause: illegal config
    _bFault := TRUE;                           // 标志与码位配对（R45） / Flag paired with code
END_IF

(* —— 段 3：落料超时与满 bin 换道（判据当拍量；下标写前钳制） —— *)
IF (NOT _bFault) AND tonDrop.Q THEN            // 落料超时 / Drop timeout
    _uFault := 16#0005_03A1;
    _eCause := E_DL_OcvCause.eDropTmo;         // 归因：落料超时 / Cause: drop timeout
    _bFault := TRUE;
END_IF
IF (NOT _bFault) AND (_nGrade >= 1) AND (_nGrade <= 4)
   AND (_anBinUsed[_nGrade] >= nBinCap) AND (NOT bBinCleared) THEN   // 目标 bin 已满且未清空 / Target bin full
    _uFault := 16#0005_03A1;
    _eCause := E_DL_OcvCause.eBinFull;         // 归因：满 bin 换道 / Cause: bin full
    _bFault := TRUE;
END_IF

(* —— 段 4：故障解除式（R240；全当拍量）：rtReset.Q / NOT _bCfgBad / NOT tonDrop.Q / bBinCleared —— *)
IF rtReset.Q AND (NOT _bCfgBad) AND (NOT tonDrop.Q) AND bBinCleared THEN
    _bFault := FALSE;                          // 清故障锁存位（锁存量） / Clear fault latch
    _uFault := 16#0000_0000;                   // 清故障锁存码（锁存量） / Clear fault code
    _eCause := E_DL_OcvCause.eNone;            // 清成因（锁存量） / Clear cause
END_IF

(* —— 段 4A：故障锁存相位迁移闸 —— *)
IF _bFault AND (_eState <> E_DL_OcvState.eFault) THEN
    _eState := E_DL_OcvState.eFault;           // 锁存即入故障相 / Latch enters fault phase
END_IF

(* —— 段 5：相位机（CASE 全覆盖 + ELSE 兜底） —— *)
CASE _eState OF

E_DL_OcvState.eIdle:
    IF bStart AND (NOT _bFault) THEN           // 启动条件 / Start gate
        _eState := E_DL_OcvState.eClassify;    // 进档位判定相 / Enter classification
    END_IF

E_DL_OcvState.eClassify:
    IF (_nGrade >= 1) AND (_nGrade <= 4) THEN  // 出口 1：档位有效（下标已钳制） / Valid grade
        _eState := E_DL_OcvState.eDispatch;    // 进落料相 / Enter dispatch
    ELSIF NOT bStart THEN                      // 出口 2：撤启动（R98 双出口） / Start released
        _eState := E_DL_OcvState.eIdle;
    END_IF

E_DL_OcvState.eDispatch:
    IF tonDrop.Q THEN                          // 落料到时 / Drop elapsed
        IF (_nGrade >= 1) AND (_nGrade <= 4) AND (NOT (_anBinUsed[_nGrade] >= nBinCap)) THEN
            _anBinUsed[_nGrade] := _anBinUsed[_nGrade] + 1;   // 计数递增（钳制下标 + 容量复核） / Increment with clamped index
        END_IF
        _uInfo := 16#0005_04C9;                // 信息级：单件分选完成沿 / Info: piece sorted edge
        _eState := E_DL_OcvState.eDone;        // 进完成相 / Enter done
    ELSIF NOT bStart THEN                      // 撤启动：中止 / Abort
        _eState := E_DL_OcvState.eIdle;
    END_IF

E_DL_OcvState.eDone:
    IF NOT bStart THEN                         // 撤启动回空闲 / Start released returns idle
        _eState := E_DL_OcvState.eIdle;
    END_IF

E_DL_OcvState.eFault:
    ;                                          // 故障相：仅段 4 复位沿可迁出 / Only reset exits

ELSE
    _uFault := 16#0005_03A1;                   // 故障级：非法相位兜底（归并总码） / Illegal phase fallback
    _eCause := E_DL_OcvCause.eCfgIllegal;      // 归因：相位非法归并组态 / Cause: phase illegal
    _bFault := TRUE;
    _eState := E_DL_OcvState.eFault;           // 强制回故障相 / Force fault phase

END_CASE

(* —— 段 6：出口单点映射（名实同源；锁存码回放） —— *)
nGrade := _nGrade;                             // 档位出口 / Grade outlet
anBinUsed[1] := _anBinUsed[1];                 // 1 档计数映射 / Grade 1 usage
anBinUsed[2] := _anBinUsed[2];                 // 2 档计数映射 / Grade 2 usage
anBinUsed[3] := _anBinUsed[3];                 // 3 档计数映射 / Grade 3 usage
anBinUsed[4] := _anBinUsed[4];                 // 4 档计数映射 / Grade 4 usage
bBinFull := (_nGrade >= 1) AND (_nGrade <= 4) AND (_anBinUsed[_nGrade] >= nBinCap);  // 满 bin 镜像 / Bin full mirror
bCycleDone := (_eState = E_DL_OcvState.eDone);// 完成标志 / Done flag
IF _bFault THEN
    nErrId := _uFault;                         // 故障锁存码回放 / Replay latched code
ELSE
    nErrId := _uInfo;                          // 信息码 / Transient info
END_IF
bError := _bFault;                             // 故障标志同源 / Flag from latch
eState := _eState;                             // 状态出口 / State outlet
eCause := _eCause;                             // 成因出口 / Cause outlet

END_FUNCTION_BLOCK

(* ---- FB_DL_CellSortingBin.st ---- *)
(*==============================================================================
 * 组件名称 (Component)  : FB_DL_CellSortingBin
 * 所属子库 (Sublibrary) : DL_Process
 * 当前版本 (Version)    : 1.0.0
 * 兼容性   (Platform)   : CODESYS 3.5+ / TwinCAT 3 / 汇川 InoProShop / 施耐德 Machine Expert
 *                         仅依赖 Standard.library（R_TRIG），零厂商私有库
 * 功能描述 (Function)   : 电池片分选落料 + 料仓满溢调度。
 *                           ① 档位→料仓映射：anGradeMap[nGrade − 1] 给出目标仓号，−1 表示该档
 *                              "不落料"（工艺上存在 NG 档直接走废料带、不进分选仓的情形）。
 *                           ② 满溢调度：目标仓已满（anBinCount ≥ anBinCapacity）时**不丢片**，
 *                              自动旁路到备仓 nBackupBin，并置 bOverflowBypass 锁存告警
 *                              （旁路是被动降级，必须让维护看见；悄悄丢片是最坏结果）。
 *                           ③ 双满兜底：目标仓与备仓同时满 → bNoBin 锁存故障、不落料、
 *                              由上层停机或切换收料框（本件不擅自选第三个仓——仓序属产线配置，
 *                              不是算法可以推断的）。
 *                           ④ 计数在**成功落料后**自增（inc-place 写回调用方的 anBinCount），
 *                              杜绝"先计数后落料"导致的仓位数虚高。
 * 接口     (Interface)  : 输入 nGrade 当前档位（1..8）、bDropCmd 落料命令（上升沿执行）、
 *                         anBinCount 各仓当前计数（VAR_IN_OUT，成功落料后自增）、
 *                         anBinCapacity 各仓容量（配置）、anGradeMap 档位到料仓映射（配置，−1 不落）、
 *                         nBackupBin 备仓号、bReset 复位；输出 nTargetBin 目标仓（−1 无）、
 *                         bDrop 落料脉冲（单拍）、bOverflowBypass 旁路告警（锁存）、
 *                         bNoBin 无可用仓（锁存）、bGradeUnmapped 该档不落料（当拍量）、
 *                         eState / eCause / bError。
 * 边界     (Boundary)   : ① **属主边界（写死）：本件只做"档位到仓号的选择与满溢旁路"，
 *                         不驱动气缸/翻转机构、不做到位确认**。执行机构动作与到位联锁属
 *                         落料执行 POU（可复用 `I_DL_Cylinder` 族）；本件只出目标仓号与落料脉冲。
 *                         ② 组态闸：nGrade < 1 或 > 8（越映射表边界）、nBackupBin 越 0..3、
 *                         任一 anBinCapacity[i] <= 0、映射表值 > 3（越仓边界）或 < −1、
 *                         映射表指向的仓不存在 → 故障锁存，落料脉冲不出（宁可不落，不可乱落）。
 *                         ③ 4 仓定长（ARRAY[0..3]）、8 档定长（ARRAY[0..7]）：容量写死在类型里，
 *                         改仓数须改类型定义，不允许"运行期可变长度"（那会越界）。
 *                         ④ 单枚 R_TRIG（bDropCmd）+ 单枚 R_TRIG（bReset）段 0 无条件周期刷新；
 *                         无 TON，故无跨相复位风险。
 *                         ⑤ 故障相与旁路锁存迁出唯一路径 = bReset 上升沿（R228B）。
 *                         ⑥ 零全局耦合（无 GVL / 无 VAR_EXTERNAL / 无物理地址）。
 * 分工声明 (Scope)      : 与 `FB_DL_Cylinder` 族（执行机构）分工——本件是**调度/记账**件，
 *                         输出仓号与脉冲；执行件负责把片真送进仓。二者不可混写在一个 FB 里，
 *                         否则换执行机构时要重测记账逻辑。
 * 来源标签 (Source Tag) : ROADMAP B 类（光伏电池片分选落料，自研 clean-room，无外源代码）
 * 解除式   (Release)    : bReset 上升沿 ∧ 组态合法 → 清 bNoBin / bOverflowBypass 锁存。
 *                         自证可满足：清仓（计数减少）或复位后即解除，无恒假因子。
 * 码表     (Codes)      : 本件不占用任何全局数字码位。出口为 INT 仓号 + BOOL 组 + ENUM
 *                         （eState / eCause）；数字码位待主控收口阶段统一派号。
 * 红线自检 (Redline)    : R1 ✓ 零 GVL/VAR_EXTERNAL ｜ R2 ✓ 零 %I/%Q/%M ｜ R3 ✓ 纯 IEC 61131-3
 *                         R4 ✓ 数组边界闸 + 映射值域闸 + 容量非正闸 ｜ R5 ✓ 声明逐行同行双语注释
 *                         R6 ✓ ENUM+CASE 含 ELSE ｜ R7 ✓ R_TRIG 段 0 无条件刷新
 * 修订历史 (Revision)   : 2026-11-19  v1.0.0  R46 首版（批次 3 · 序号 14）
 *==============================================================================*)

TYPE E_DL_CsbState :
(
    eIdle  := 0,    // 等待落料命令 / Awaiting a drop command
    eRun   := 10,   // 正常落料运行相 / Normal dropping
    eBypass:= 20,   // 满溢旁路相（走备仓，告警保持） / Overflow bypass phase
    eFault := 90    // 无可用仓/组态故障相 / No-bin or configuration fault
);
END_TYPE

TYPE E_DL_CsbCause :
(
    eNone        := 0,   // 无异常 / No anomaly
    eCfgIllegal  := 1,   // 组态非法（映射/容量/备仓越界） / Illegal configuration
    eOverflow    := 2,   // 目标仓满溢，已旁路到备仓 / Target bin full, bypassed to the backup bin
    eNoBin       := 3,   // 目标仓与备仓同时满，无可用仓 / Target and backup both full
    eGradeUnmapped:= 4,  // 该档不落料（映射为 −1） / Grade intentionally not dropped
    ePhaseBad    := 5    // 非法相位兜底 / Illegal phase fallback
);
END_TYPE

FUNCTION_BLOCK FB_DL_CellSortingBin
VAR_IN_OUT
    anBinCount : ARRAY[0..3] OF DINT;       // 各仓当前计数（成功落料后本件自增） [片] / Bin counts, incremented by this unit on success [pcs]
END_VAR
VAR_INPUT
    nGrade        : INT := 1;               // 当前档位，域 1..8 / Present grade, 1..8
    bDropCmd      : BOOL := FALSE;          // 落料命令，上升沿执行一次 [-] / Drop command, acts once per rising edge
    anBinCapacity : ARRAY[0..3] OF DINT;    // 各仓容量（配置），每项域 > 0 [片] / Bin capacities, each > 0 [pcs]
    anGradeMap    : ARRAY[0..7] OF INT;     // 档位到仓映射（配置），值域 −1 或 0..3 [-] / Grade-to-bin map, -1 or 0..3
    nBackupBin    : INT := 3;               // 备仓号，域 0..3 / Backup bin index, 0..3
    bReset        : BOOL := FALSE;          // 复位，上升沿清旁路与无仓锁存 [-] / Reset, rising edge clears latches
END_VAR
VAR_OUTPUT
    nTargetBin      : INT;                  // 本拍目标仓号，−1 表示无 / Target bin this scan, -1 means none
    bDrop           : BOOL;                 // 落料脉冲（单拍） [-] / Drop pulse, single scan
    bOverflowBypass : BOOL;                 // 满溢旁路告警（锁存） [-] / Overflow bypass alarm, latched
    bNoBin          : BOOL;                 // 无可用仓（锁存故障） [-] / No available bin, latched fault
    bGradeUnmapped  : BOOL;                 // 该档不落料（当拍量，非故障） [-] / Grade not dropped, per scan, not a fault
    eState          : E_DL_CsbState;        // 状态出口 [-] / State outlet
    eCause          : E_DL_CsbCause;        // 成因出口（R190 归因唯一） [-] / Cause outlet
    bError          : BOOL;                 // 故障标志（无仓/组态非法；旁路不算故障） [-] / Error flag, bypass is not a fault
END_VAR
VAR
    _eState   : E_DL_CsbState := E_DL_CsbState.eIdle;    // 内部相位（CASE 唯一写入目标） / Internal phase
    _eCause   : E_DL_CsbCause := E_DL_CsbCause.eNone;    // 成因锁存量 / Latched cause
    rtDrop    : R_TRIG;                 // 落料命令沿实例，段 0 无条件调用 / Drop edge instance
    rtReset   : R_TRIG;                 // 复位沿实例，段 0 无条件调用 / Reset edge instance
    _bBypass  : BOOL;                   // 旁路告警锁存位（锁存量） / Latched bypass alarm
    _bNoBin   : BOOL;                   // 无可用仓锁存位（锁存量） / Latched no-bin fault
    _bCfgBad  : BOOL;                   // 组态非法当拍量 [-] / Illegal configuration this scan
    _bMapBad  : BOOL;                   // 映射表非法当拍量 [-] / Illegal map this scan
    _nBin     : INT;                    // 映射得到的目标仓号中间量 [-] / Mapped target bin intermediate
    _nMapIdx  : INT;                    // 映射查表索引（已钳位） [-] / Clamped map index
    _i        : INT;                    // 遍历索引 / Loop index
END_VAR
VAR CONSTANT
    DL_CSB_BINMAX : INT := 3;           // 仓号上界（与 ARRAY[0..3] 一致） [仓] / Bin index bound matching the array
    DL_CSB_GRDMAX : INT := 8;           // 档位上界（与 ARRAY[0..7] 一致） [档] / Grade bound matching the array
    DL_CSB_NOBIN  : INT := -1;          // 无目标仓哨兵值 [-] / Sentinel for "no target bin"
END_VAR

(* —— 段 0：组态闸派生 + 两沿实例无条件周期刷新 —— *)
_bMapBad := FALSE;                                          // 映射非法初值 / Map-illegal initial value
FOR _i := 0 TO DL_CSB_GRDMAX - 1 DO
    IF (anGradeMap[_i] > DL_CSB_BINMAX) OR (anGradeMap[_i] < DL_CSB_NOBIN) THEN
        _bMapBad := TRUE;                                   // 映射值越界（> 3 或 < −1） / Map value out of range
    END_IF
END_FOR
FOR _i := 0 TO DL_CSB_BINMAX DO
    IF anBinCapacity[_i] <= 0 THEN
        _bMapBad := TRUE;                                   // 容量非正（永不装满或立即装满，皆病态） / Non-positive capacity is degenerate
    END_IF
END_FOR
_bCfgBad := _bMapBad
        OR (nBackupBin < 0) OR (nBackupBin > DL_CSB_BINMAX)   // 备仓号越界 / Backup index out of range
        OR (nGrade < 1) OR (nGrade > DL_CSB_GRDMAX);          // 档位越映射表边界 / Grade out of the map bounds
rtDrop(CLK := bDropCmd);                                    // 落料沿，每拍必调（R228A） / Drop edge, every scan
rtReset(CLK := bReset);                                     // 复位沿，每拍必调 / Reset edge, every scan

(* —— 段 1：单拍量预清零（锁存量 _bBypass / _bNoBin / _eCause 不入清单，R107） —— *)
nTargetBin     := DL_CSB_NOBIN;     // 目标仓缺省无 / Target bin defaults to none
bDrop          := FALSE;            // 落料脉冲每拍预清 / Drop pulse preset
bOverflowBypass:= FALSE;            // 旁路出口每拍预清 / Bypass outlet preset
bNoBin         := FALSE;            // 无仓出口每拍预清 / No-bin outlet preset
bGradeUnmapped := FALSE;            // 不落料标志每拍预清 / Unmapped flag preset
bError         := FALSE;            // 故障标志每拍预清（R45 配对） / Error flag preset

(* —— 段 2：复位沿 + 组态闸 —— *)
IF rtReset.Q THEN
    _bBypass := FALSE;                                  // 清旁路告警锁存 / Clear the bypass alarm
    _bNoBin  := FALSE;                                  // 清无仓锁存 / Clear the no-bin latch
    _eCause  := E_DL_CsbCause.eNone;                    // 清成因 / Clear cause
    IF _eState = E_DL_CsbState.eFault THEN
        _eState := E_DL_CsbState.eIdle;                 // 故障相迁出（R228B） / Leave fault phase
    END_IF
    IF _eState = E_DL_CsbState.eBypass THEN
        _eState := E_DL_CsbState.eRun;                  // 旁路相迁出（第二条可迁出路径） / Leave bypass phase, second exit path
    END_IF
END_IF
IF _bCfgBad THEN
    _eState := E_DL_CsbState.eFault;                    // 入故障相 / Enter fault phase
    _eCause := E_DL_CsbCause.eCfgIllegal;               // 归因：组态非法 / Cause: illegal configuration
END_IF

(* —— 段 3：落料调度（命令沿 + 组态合法；单点写入锁存与计数） —— *)
IF rtDrop.Q AND (NOT _bCfgBad) THEN
    _nMapIdx := nGrade - 1;                             // 映射查表索引（段 0 已闸 1..8） / Map index, grade bounds already gated
    IF _nMapIdx < 0 THEN
        _nMapIdx := 0;                                  // 下界钳（双保险） / Lower clamp, second guard
    END_IF
    IF _nMapIdx > DL_CSB_GRDMAX - 1 THEN
        _nMapIdx := DL_CSB_GRDMAX - 1;                  // 上界钳（双保险） / Upper clamp, second guard
    END_IF
    _nBin := anGradeMap[_nMapIdx];                      // 目标仓号 / Mapped target bin
    IF _nBin = DL_CSB_NOBIN THEN
        bGradeUnmapped := TRUE;                         // 该档不落料（工艺意图，非故障） / Grade intentionally not dropped
        _eCause := E_DL_CsbCause.eGradeUnmapped;        // 成因：映射为不落料 / Cause: mapped to no-drop
    ELSE
        IF anBinCount[_nBin] < anBinCapacity[_nBin] THEN
            nTargetBin := _nBin;                        // 目标仓有余量，正常落 / Target bin has room
            anBinCount[_nBin] := anBinCount[_nBin] + 1; // 成功落料后计数（先判满后自增） / Increment only after a successful drop
            bDrop := TRUE;                              // 落料脉冲 / Drop pulse
            IF _eState = E_DL_CsbState.eIdle THEN
                _eState := E_DL_CsbState.eRun;          // 首次落料入运行相 / First drop enters run
            END_IF
        ELSIF anBinCount[nBackupBin] < anBinCapacity[nBackupBin] THEN
            nTargetBin := nBackupBin;                   // 旁路到备仓 / Bypass to the backup bin
            anBinCount[nBackupBin] := anBinCount[nBackupBin] + 1;   // 备仓计数自增 / Increment the backup bin
            bDrop := TRUE;                              // 落料脉冲 / Drop pulse
            _bBypass := TRUE;                           // 旁路告警锁存（被动降级必须可见） / Latch the bypass alarm
            _eCause := E_DL_CsbCause.eOverflow;         // 成因：满溢旁路 / Cause: overflow bypass
            _eState := E_DL_CsbState.eBypass;           // 入旁路相 / Enter the bypass phase
        ELSE
            nTargetBin := DL_CSB_NOBIN;                 // 双满：无可用仓 / Both full: no available bin
            _bNoBin := TRUE;                            // 无仓锁存故障 / Latch the no-bin fault
            _eCause := E_DL_CsbCause.eNoBin;            // 成因：无可用仓 / Cause: no available bin
            _eState := E_DL_CsbState.eFault;            // 入故障相 / Enter the fault phase
        END_IF
    END_IF
END_IF

(* —— 段 4：锁存相位迁移闸（无仓故障必须停在故障相，旁路必须停在旁路相） —— *)
IF _bNoBin AND (_eState <> E_DL_CsbState.eFault) THEN
    _eState := E_DL_CsbState.eFault;                    // 无仓锁存即入故障相 / No-bin latch enters fault
END_IF

(* —— 段 5：相位机（ENUM 全成员显式标签 + ELSE 兜底，R128） —— *)
CASE _eState OF

E_DL_CsbState.eIdle:
    IF _bCfgBad THEN                                    // 出口 1：组态非法 / Illegal configuration
        _eState := E_DL_CsbState.eFault;
    ELSIF rtDrop.Q AND (NOT _bCfgBad) THEN              // 出口 2：已有落料动作 / A drop has been dispatched
        _eState := E_DL_CsbState.eRun;
    END_IF

E_DL_CsbState.eRun:
    IF _bCfgBad OR _bNoBin THEN                         // 出口 1：故障（组态或无仓） / Fault, config or no-bin
        _eState := E_DL_CsbState.eFault;
    ELSIF _bBypass THEN                                 // 出口 2：发生过满溢旁路 / An overflow bypass occurred
        _eState := E_DL_CsbState.eBypass;
    END_IF

E_DL_CsbState.eBypass:
    IF _bNoBin THEN                                     // 出口 1：旁路后仍双满 / Both full even after bypass
        _eState := E_DL_CsbState.eFault;
    ELSIF _bBypass = FALSE THEN                         // 出口 2：旁路告警被复位清除 / Bypass alarm cleared by reset
        _eState := E_DL_CsbState.eRun;
    END_IF

E_DL_CsbState.eFault:
    ;                                                   // 故障相：仅段 2 复位沿可迁出 / Only the reset edge leaves this phase

ELSE
    _eCause := E_DL_CsbCause.ePhaseBad;                 // 归因：非法相位 / Cause: illegal phase
    _eState := E_DL_CsbState.eFault;                    // 强拉故障相 / Force the fault phase
    bError  := TRUE;                                    // 故障标志 / Error flag

END_CASE

(* —— 段 6：出口单点映射（名实双出口，R191；旁路是告警不是故障，此处写死分级） —— *)
bOverflowBypass := _bBypass;                            // 旁路告警与锁存同源 / Bypass alarm from latch
bNoBin          := _bNoBin;                             // 无仓与锁存同源 / No-bin from latch
bError          := _bNoBin OR _bCfgBad;                 // 故障标志：无仓或组态非法（旁路不计入故障级） / Error: no-bin or illegal config, bypass excluded
eState          := _eState;                             // 状态出口 / State outlet
eCause          := _eCause;                             // 成因出口 / Cause outlet

END_FUNCTION_BLOCK

(* ---- FB_DL_CentrifugeSpinSeq.st ---- *)
(*
  道莅工业代码库 | DL_Process | FB_DL_CentrifugeSpinSeq
  版本: 1.0.0 | 日期: 2026-11-23 | 轮次: R75
  开源溯源: self-cleanroom（无外部来源；行业池·分离设备通用语义，零代码行复制）
  功能: 离心机升速-恒速-降速三段序列，含临界转速快跳段（给定直接跳过临界带，
        实测转速越带上沿后恢复斜坡）与不平衡/开盖/转速非有限三路停机闸（跳闸锁存）。
  兼容性: CODESYS 3.5 / TwinCAT 3 / 汇川 InoProShop；仅依赖标准 TON / R_TRIG / LIMIT，零厂商私有库
  接口: 输入启动/盖开关/实测转速/目标转速/临界带/升降斜率/周期/不平衡信号/复位；
        输出 fSpRef [rpm]/bDriveEn/bBrakeOut/bAtSpeed/eState/eCause/bError/nErrId。
  码表: 16#0005_03BA 故障级：离心机跳闸总码（锁存至复位沿，归由 eCause）
        码段说明：0005 段故障子带 03xx，槽位经全库实扫空闲。
  边界: ① 快跳段：给定值在临界带内不给斜坡、直接跳带上沿（fCritHi），
        实测转速 >= fCritHi - 容差 后回 eAccel 续斜坡（避开共振驻留）；
        ② 不平衡经 tUnbalDelay 去抖确认跳闸；开盖/转速 NaN 即时跳闸；
        ③ 跳闸相：驱动禁止 + 制动输出，唯一解除路径 = bReset 上升沿 ∧
        组态合法 ∧ 盖已关；
        ④ 斜坡积分上限：MIN(fSpeedSp)；降速下限钳 0；
        ⑤ TON/R_TRIG 段 0 无条件周期刷新；⑥ 零全局耦合。
  邻件比对: registry 扫查 centrifuge 零命中（R75 §3 留痕），无属主。
  修订历史: 2026-11-23 v1.0.0 R75 首版（复杂件批 B2 · C08）
*)

TYPE E_DL_CssState :
(
    eIdle  := 0,   // 待机（给定钳零，驱动禁止） | Idle, ref zero, drive off
    eAccel := 10,  // 斜坡升速 | Ramped acceleration
    eCrit  := 20,  // 临界转速快跳段 | Critical band fast jump
    eRun   := 30,  // 恒速运行 | Constant speed run
    eDecel := 40,  // 斜坡降速 | Ramped deceleration
    eTrip  := 90   // 跳闸锁存相（驱动禁止+制动） | Trip latch phase
);
END_TYPE

TYPE E_DL_CssCause :
(
    eNone          := 0,  // 无故障 | No cause
    eCfgIllegal    := 1,  // 组态非法 | Illegal configuration
    eUnbalance     := 2,  // 不平衡超限（去抖确认） | Unbalance confirmed by debounce
    eLidOpen       := 3,  // 运转中开盖 | Lid opened in motion
    eSensNonFinite := 4   // 转速反馈非有限 | Speed feedback non-finite
);
END_TYPE

FUNCTION_BLOCK FB_DL_CentrifugeSpinSeq
VAR_INPUT
    bStartCmd    : BOOL := FALSE;    // 启动命令（电平）[-] | Start command level
    bLidClosed   : BOOL := TRUE;     // 盖已关（安全联锁）[-] | Lid closed interlock
    fSpeedAct    : REAL := 0.0;      // 实测转速 [rpm] | Speed feedback actual
    fSpeedSp     : REAL := 3000.0;   // 目标转速，域 > fCritHi [rpm] | Target speed setpoint
    fCritLo      : REAL := 800.0;    // 临界转速带下沿，域 < 上沿 [rpm] | Critical band lower edge
    fCritHi      : REAL := 1100.0;   // 临界转速带上沿，域 < 目标转速 [rpm] | Critical band upper edge
    fRampUp      : REAL := 100.0;    // 升速斜率，域 > 0 [rpm/s] | Ramp-up rate
    fRampDn      : REAL := 200.0;    // 降速斜率，域 > 0 [rpm/s] | Ramp-down rate
    fDtSec       : REAL := 0.01;     // 序列周期，域 (0, 1] [s] | Sequence cycle time
    fAtSpeedTol  : REAL := 30.0;     // 到速容差，域 > 0 [rpm] | At-speed tolerance
    fStopThresh  : REAL := 10.0;     // 停转判据阈值，域 > 0 [rpm] | Stopped threshold
    tUnbalDelay  : TIME := T#2S;     // 不平衡确认延时，域 > T#0S | Unbalance confirm delay
    bUnbalHigh   : BOOL := FALSE;    // 不平衡检测输入（电平）[-] | Unbalance detection level
    bReset       : BOOL := FALSE;    // 复位命令，上升沿清跳闸 [-] | Reset command, rising edge
END_VAR
VAR_OUTPUT
    fSpRef    : REAL;               // 转速给定出口 [rpm] | Speed reference outlet
    bDriveEn  : BOOL;               // 驱动使能出口 [-] | Drive enable outlet
    bBrakeOut : BOOL;               // 制动输出出口 [-] | Brake output outlet
    bAtSpeed  : BOOL;               // 到速判据出口 [-] | At-speed outlet
    eState    : E_DL_CssState;      // 状态出口 | State outlet
    eCause    : E_DL_CssCause;      // 跳闸成因出口 | Trip cause outlet
    bError    : BOOL;               // 故障锁存标志 [-] | Fault latch flag
    nErrId    : UDINT;              // 事件码，0 = 无事件 | Event code, 0 = none
END_VAR
VAR
    _eState  : E_DL_CssState := E_DL_CssState.eIdle;   // 内部状态（CASE 唯一写入目标） | Internal state
    _eCause  : E_DL_CssCause := E_DL_CssCause.eNone;   // 成因锁存 | Latched cause
    _bFault  : BOOL;            // 故障锁存位 | Fault latch bit
    _fSpRef  : REAL := 0.0;     // 给定积分内部镜像 [rpm] | Reference ramp internal mirror
    _bCfgBad : BOOL;            // 组态非法当拍量 [-] | Illegal configuration
    _bSensBad: BOOL;            // 转速反馈非有限当拍量 [-] | Speed feedback non-finite
    rtStart  : R_TRIG;          // 启动沿实例，段 0 无条件刷新 | Start edge instance
    rtReset  : R_TRIG;          // 复位沿实例，段 0 无条件刷新 | Reset edge instance
    tonUnbal : TON;             // 不平衡去抖计时，段 0 无条件刷新 | Unbalance debounce timer
END_VAR
VAR CONSTANT
    DL_CSS_EPS : REAL := 1.0;       // 快跳越带容差 [rpm] | Jump exit tolerance
    DL_CSS_ERR : UDINT := 16#0005_03BA;  // 跳闸故障码 | Trip fault code
END_VAR

(* —— 段 0：当拍量派生 + 定时器与沿实例无条件周期刷新（R7 红线） —— *)
_bSensBad := (fSpeedAct <> fSpeedAct);                                      // 转速反馈 NaN 自反判 / Speed NaN self-reflex check
_bCfgBad := (fCritLo >= fCritHi) OR (fSpeedSp <= fCritHi) OR (fRampUp <= 0.0)
         OR (fRampDn <= 0.0) OR (fDtSec <= 0.0) OR (fDtSec > 1.0)
         OR (fAtSpeedTol <= 0.0) OR (fStopThresh <= 0.0)
         OR (fSpeedSp <> fSpeedSp) OR (fCritLo <> fCritLo) OR (fCritHi <> fCritHi);  // 组态域闸（含组态量非有限）/ Configuration gate
rtStart(CLK := bStartCmd);                                                  // 启动沿每拍必调 / Start edge every scan
rtReset(CLK := bReset);                                                     // 复位沿每拍必调 / Reset edge every scan
tonUnbal(IN := bUnbalHigh AND ((_eState = E_DL_CssState.eAccel)
         OR (_eState = E_DL_CssState.eCrit) OR (_eState = E_DL_CssState.eRun)), PT := tUnbalDelay); // 不平衡去抖 IN 挂运转相 ∧ 信号 / Debounce gated by motion and signal

(* —— 段 1：复位沿 + 组态域闸 —— *)
IF rtReset.Q AND (NOT _bCfgBad) AND bLidClosed THEN                         // 复位沿且组态合法且盖已关 / Reset with legal config and lid closed
    _bFault := FALSE;                                                       // 清故障锁存位 / Clear fault latch
    _eCause := E_DL_CssCause.eNone;                                         // 清成因 / Clear cause
    IF _eState = E_DL_CssState.eTrip THEN
        _eState := E_DL_CssState.eIdle;                                     // 跳闸相迁出唯一路径 / Sole trip exit
    END_IF
END_IF
IF _bCfgBad THEN                                                            // 组态域闸 / Configuration gate
    _bFault := TRUE;
    _eCause := E_DL_CssCause.eCfgIllegal;                                   // 归因组态 / Cause: config
END_IF

(* —— 段 2：运转相即时跳闸源（开盖 / 转速非有限） —— *)
IF (NOT _bFault) AND ((_eState = E_DL_CssState.eAccel)
    OR (_eState = E_DL_CssState.eCrit) OR (_eState = E_DL_CssState.eRun)) THEN
    IF NOT bLidClosed THEN
        _bFault := TRUE;                                                    // 运转中开盖即时跳闸 / Lid open in motion, immediate trip
        _eCause := E_DL_CssCause.eLidOpen;                                  // 归因开盖 / Cause: lid open
    ELSIF _bSensBad THEN
        _bFault := TRUE;                                                    // 转速反馈丢失即时跳闸 / Speed feedback loss trip
        _eCause := E_DL_CssCause.eSensNonFinite;                            // 归因反馈 / Cause: feedback
    END_IF
END_IF

(* —— 段 3：不平衡去抖跳闸（三运转相共用一码，R190 归因唯一） —— *)
IF (NOT _bFault) AND tonUnbal.Q THEN
    _bFault := TRUE;                                                        // 不平衡跳闸锁存 / Unbalance trip latch
    _eCause := E_DL_CssCause.eUnbalance;                                    // 归因不平衡 / Cause: unbalance
END_IF

(* —— 段 4：状态机（ENUM + CASE，ELSE 兜底） —— *)
CASE _eState OF

E_DL_CssState.eIdle:
    _fSpRef := 0.0;                                                         // 待机给定钳零 / Idle ref zero
    IF rtStart.Q AND bLidClosed AND (NOT _bFault) THEN
        _fSpRef := 0.0;                                                     // 启动给定从零起 ramp / Start ramp from zero
        _eState := E_DL_CssState.eAccel;                                    // 进入升速段 / Enter accel
    END_IF

E_DL_CssState.eAccel:
    _fSpRef := _fSpRef + fRampUp * fDtSec;                                  // 斜坡升速积分 [rpm] / Ramp-up integration
    _fSpRef := LIMIT(0.0, _fSpRef, fSpeedSp);                               // 给定钳 [0, fSpeedSp] / Reference clamp
    IF _fSpRef >= fCritLo THEN
        _eState := E_DL_CssState.eCrit;                                     // 给定达临界带下沿转快跳 / Ref at band lower edge, jump
    ELSIF _fSpRef >= fSpeedSp THEN
        _eState := E_DL_CssState.eRun;                                      // 无临界带穿越直达恒速（组态已闸 fSpeedSp > fCritHi，防御分支） / Direct to run, defensive
    ELSIF (NOT bStartCmd) THEN
        _eState := E_DL_CssState.eDecel;                                    // 启动命令撤转降速 / Start released, decel
    END_IF

E_DL_CssState.eCrit:
    _fSpRef := fCritHi;                                                     // 快跳段：给定直接跳带上沿（边界①）/ Fast jump to upper edge
    IF fSpeedAct >= (fCritHi - DL_CSS_EPS) THEN
        _eState := E_DL_CssState.eAccel;                                    // 实测越带上沿回斜坡续升 / Feedback past band, resume ramp
    ELSIF (NOT bStartCmd) THEN
        _eState := E_DL_CssState.eDecel;                                    // 快跳段内命令撤转降速 / Start released in jump, decel
    END_IF

E_DL_CssState.eRun:
    _fSpRef := fSpeedSp;                                                    // 恒速段给定锁目标 / Run ref at target
    IF (NOT bStartCmd) THEN
        _eState := E_DL_CssState.eDecel;                                    // 命令撤转降速 / Start released, decel
    END_IF

E_DL_CssState.eDecel:
    _fSpRef := _fSpRef - fRampDn * fDtSec;                                  // 斜坡降速积分 [rpm] / Ramp-down integration
    IF _fSpRef < 0.0 THEN
        _fSpRef := 0.0;                                                     // 给定下限钳零 / Ref clamp zero
    END_IF
    IF (_fSpRef <= 0.0) AND (fSpeedAct < fStopThresh) THEN
        _eState := E_DL_CssState.eIdle;                                     // 给定归零且实测停转回待机 / Ref zero and stopped, idle
    END_IF

E_DL_CssState.eTrip:
    _fSpRef := 0.0;                                                         // 跳闸给定钳零 / Trip ref zero
    ;                                                                       // 仅段 1 复位沿可迁出 / Only reset edge leaves

ELSE
    _bFault := TRUE;                                                        // 非法状态兜底（R6）/ Illegal state fallback
    _eCause := E_DL_CssCause.eCfgIllegal;                                   // 归因归并组态 / Cause folded to config
    _eState := E_DL_CssState.eTrip;

END_CASE

(* —— 段 5：出口单点映射（名实同源；锁存码回放） —— *)
fSpRef := _fSpRef;                                                          // 给定出口 [rpm] / Reference outlet
bDriveEn := (_eState = E_DL_CssState.eAccel) OR (_eState = E_DL_CssState.eCrit)
         OR (_eState = E_DL_CssState.eRun) OR (_eState = E_DL_CssState.eDecel);  // 驱动使能四运转相 / Drive enable in motion states
bBrakeOut := (_eState = E_DL_CssState.eDecel) OR (_eState = E_DL_CssState.eTrip);  // 制动输出降速/跳闸相 / Brake in decel and trip
bAtSpeed := (_eState = E_DL_CssState.eRun) AND (fSpeedAct >= (fSpeedSp - fAtSpeedTol));  // 到速判据 / At-speed judgement
eState := _eState;                                                          // 状态出口 / State outlet
eCause := _eCause;                                                          // 成因出口 / Cause outlet
bError := _bFault;                                                          // 故障标志同源 / Error flag from latch
IF _bFault THEN
    nErrId := DL_CSS_ERR;                                                   // 跳闸锁存码回放 / Replay latched trip code
ELSE
    nErrId := 16#0000_0000;                                                 // 无事件 / No event
END_IF

END_FUNCTION_BLOCK

(* ---- FB_DL_ChamberLeakRate.st ---- *)
(*==============================================================================
 * 组件名称 (Component)  : FB_DL_ChamberLeakRate
 * 所属子库 (Sublibrary) : DL_Process
 * 前缀     (Prefix)     : FB_DL_
 * 当前版本 (Version)    : 1.0.1
 * 兼容性   (Platform)   : CODESYS 3.5 / TwinCAT 3 / 汇川 InoProShop / Schneider
 *                         Machine Expert；纯 IEC 61131-3（第 3 版），
 *                         仅依赖标准库 TON / R_TRIG / ABS / MAX，零厂商方言
 * 作者     (Author)     : 道莅代码库 · PLC编程专家（R31）
 * 开源溯源 (Origin)     : 腔体压升法检漏公开工艺语义（行业池），道莅
 *                         clean-room 防御性实现，未复制任何外部源码行
 * 功能描述 (Function)   : 腔体升压率检漏件（通用压升法）。三态顺控：
 *                         稳压 → 测量 → 判定。压升率 Q = (P2 − P1)·V / tWin，
 *                         测量窗起止压强由调用方外部注入。合格判定带相对
 *                         浮点余量（1E-6 相对量），不做严格小于比较。
 * 职责边界 (Boundary)   : 与库内 EscHeLeakCheck 分工——He 背冷三段法为氦质谱
 *                         专用工艺件，本件为通用压升法单窗判定件，
 *                         二者不合并、不互替。
 * 状态机   (States)     : eIdle 待机 / eStabilize 稳压 / eMeasure 测量窗 /
 *                         eJudge 判定（单拍）/ eFault 故障锁定（CASE 带
 *                         ELSE 兜底）。
 * 码位     (Codes)      : 16#0005_0099 信息级：参数非法早退、反向压差判合格
 *                                      提示（不置 bError）
 *                         16#0005_009A 故障级：测量窗中断（测量中撤启动）
 *                         16#0005_009B 故障级：状态非法（ELSE 兜底，锁存）
 *                         16#0005_009C~009D 保留未启用（码表与实现对齐）
 * 边界防错 (Boundary)   : 1 tWin 不大于零或 V 不大于零参数非法早退（信息级）；
 *                         2 P2 < P1（反向/温降）判合格记信息码（保守侧
 *                           不误杀合格腔体）；
 *                         3 非有限全拦（x<>x 自反判加幅值界）；
 *                         4 除法分母 tWin 换算秒后强制判零；
 *                         5 故障锁存可达解除路径：重新启动沿重新受理；
 *                         6 TON/R_TRIG 实例每拍无条件刷新。
 * 修订历史 (Revision)   : 2026-11-18 v1.0.0 首版入库（R31 · 阶段三 · 序 11）
 *                         2026-11-18 v1.0.1 R31 终审修复：三处信息级码改
 *                         bInfoOne 单拍暂存，消除段 6 ELSE 同拍抹除
 *==============================================================================*)

(*------------------------------------------------------------------------------
 * 枚举: E_DL_LeakTestState（归属本功能块，同文件发布，全库唯一属主）
 *----------------------------------------------------------------------------*)
TYPE E_DL_LeakTestState :
(
    eIdle      := 0,    // 待机：未启动或已判定回位 / Idle, not started or judged
    eStabilize := 10,   // 稳压相：压力稳定等待 / Stabilize, pressure settling
    eMeasure   := 20,   // 测量相：升压测量窗计时 / Measure, leak window timing
    eJudge     := 30,   // 判定相：单拍完成判定回待机 / Judge, one-scan verdict then idle
    eFault     := 99    // 故障：测量窗中断或状态非法 / Fault, window interrupted or illegal state
);
END_TYPE

(*==============================================================================
 * 功能块: FB_DL_ChamberLeakRate
 * 调用约定: 每个扫描周期无条件调用一次；测量窗起止压强由调用方在窗口起止
 *           时刻经引脚注入（fP1 为窗起压强，fP2 为窗止压强）。
 *==============================================================================*)
FUNCTION_BLOCK FB_DL_ChamberLeakRate
VAR_INPUT
    bStart   : BOOL := FALSE;         // 启动沿（含故障态重试受理）/ Start edge, also retries from fault
    fP1      : REAL := 0.0;           // 测量窗起压强 [帕] / Window start pressure [Pa]
    fP2      : REAL := 0.0;           // 测量窗止压强 [帕] / Window end pressure [Pa]
    fV       : REAL := 1.0;           // 腔体容积 [立方米] / Chamber volume [m3]
    tWin     : TIME := T#60S;         // 测量窗时长 [毫秒] / Measurement window duration [ms]
    tStab    : TIME := T#10S;         // 稳压相时长 [毫秒]（可增引脚）/ Stabilize duration [ms], added pin
    fLeakLim : REAL := 5.0;           // 泄漏率限值 [帕立方米每秒] / Leak rate limit [Pa m3 per s]
END_VAR
VAR_OUTPUT
    fLeakRate : REAL;                 // 压升率（泄漏率）[帕立方米每秒] / Pressure rise rate [Pa m3 per s]
    bPass     : BOOL;                 // 合格标志 / Pass verdict flag
    eState    : E_DL_LeakTestState;   // 顺控当前状态 / Current sequence state
    bError    : BOOL;                 // 故障标志，与故障级码配对（R45）/ Fault flag paired with fault codes
    uErrorId  : UDINT;                // 错误码，0 = 无错 / Error code, 0 = none
END_VAR
VAR
    rTrigStart : R_TRIG;              // 启动沿检测，每拍无条件刷新 / Start edge detector, refreshed every scan
    tonPhase   : TON;                 // 相计时定时器，每拍无条件刷新 / Phase timer, refreshed every scan
    bStepRst   : BOOL;                // 相切换拍单拍断计时输入 / One-scan timer break on phase change
    tPhaseEff  : TIME;                // 本相生效计时目标 [毫秒] / Effective phase timing target [ms]
    eStatePrev : E_DL_LeakTestState;  // 上一拍状态快照 / Previous state snapshot
    bInOk      : BOOL;                // 测量输入有效性 / Measurement input validity
    bParaOk    : BOOL;                // 参数有效性 / Parameter validity
    fWinSec    : REAL;                // 测量窗秒值 [秒] / Window seconds [s]
    fRise      : REAL;                // 窗内压升 [帕] / Pressure rise over window [Pa]
    fSlack     : REAL;                // 判定浮点余量 [帕立方米每秒] / Verdict float slack [Pa m3 per s]
    uCodeLatch : UDINT;               // 故障级锁存码 / Latched fault code
    bInfoBack  : BOOL;                // 反向压差信息标志 / Reverse pressure info flag
    bInfoOne   : BOOL;                // 信息级单拍待发标志（防同拍抹除，R28 终审）/ One-scan info pending flag
    bInit      : BOOL := TRUE;        // 首扫标志 / First-scan flag
END_VAR
VAR CONSTANT
    DL_CLR_FIN  : REAL := 1.0E30;     // REAL 有限幅值判界 / REAL finiteness magnitude bound
    DL_CLR_REL  : REAL := 1.0E-6;     // 判定相对浮点余量系数 / Verdict relative slack factor
END_VAR

// ---- 段 1｜边沿与定时器实例无条件周期刷新（红线：禁入条件分支）----------------
rTrigStart(CLK := bStart);                            // 启动沿检测 / Start edge detection
tPhaseEff := tStab;                                   // 默认稳压时长 / Default stabilize duration
IF eState = eMeasure THEN
    tPhaseEff := tWin;                                // 测量相改用窗时长 / Measure phase uses window duration
END_IF
tonPhase(IN := ((eState = eStabilize) OR (eState = eMeasure)) AND (NOT bStepRst),
         PT := tPhaseEff);                            // 相计时按相取目标 / Phase timing with per-phase target

// ---- 段 2｜相切换检测（供计时器按相断输入）--------------------------------------
bStepRst := (eState <> eStatePrev) OR bInit;          // 相变化即断输入 / Phase change breaks timing input
eStatePrev := eState;                                 // 快照留痕 / Snapshot previous state
bInit := FALSE;                                       // 清首扫标志 / Clear first-scan flag

// ---- 段 3｜输入与参数有效性预判（测量相判定前复验，R42 相转换复验语义）----------
bInOk   := (fP1 = fP1) AND (fP2 = fP2) AND (ABS(fP1) < DL_CLR_FIN) AND (ABS(fP2) < DL_CLR_FIN); // 压强对有限 / Pressure pair finite
fWinSec := TIME_TO_REAL(tWin) / 1000.0;               // 窗时换算秒 [秒] / Window converted to seconds
bParaOk := (fWinSec > 0.0) AND (fV > 0.0) AND (fV = fV) AND (fV < DL_CLR_FIN); // 窗时/容积合法 / Window and volume legal

// ---- 段 4｜状态机（CASE 带 ELSE 兜底锁故障）--------------------------------------
CASE eState OF
    eIdle:
        bPass := FALSE;                               // 待机清合格标志 / Idle clears verdict
        IF rTrigStart.Q AND bParaOk THEN
            eState := eStabilize;                     // 参数合法沿进稳压 / Legal parameters, to stabilize
        ELSIF rTrigStart.Q AND (NOT bParaOk) THEN
            bInfoOne := TRUE;                         // 信息级：参数非法早退（暂存防同拍抹除）/ Info: illegal parameters, staged
        END_IF
    eStabilize:
        IF rTrigStart.Q AND (NOT bParaOk) THEN
            eState := eIdle;                          // 参数中途失配退回 / Parameters lost mid-run
            bInfoOne := TRUE;                         // 信息级：参数非法早退（暂存）/ Info: illegal parameters, staged
        ELSIF tonPhase.Q THEN
            eState := eMeasure;                       // 稳压满进测量窗 / Stabilize elapsed, to measure
            bStepRst := TRUE;                         // 单拍重载计时器入参 / One-scan timer input reload
        END_IF
    eMeasure:
        IF NOT bStart THEN
            eState := eFault;                         // 测量中撤启动即窗中断 / Start drop mid-window is interruption
            uCodeLatch := 16#0005_009A;               // 码位：测量窗中断 / Code: window interrupted
        ELSIF tonPhase.Q THEN
            eState := eJudge;                         // 窗满进判定 / Window elapsed, to judge
        END_IF
    eJudge:
        bInOk := (fP1 = fP1) AND (fP2 = fP2) AND (ABS(fP1) < DL_CLR_FIN) AND (ABS(fP2) < DL_CLR_FIN); // 判定拍复验（R42）/ Recheck at verdict scan
        bInfoBack := FALSE;                           // 反向信息先清 / Clear reverse info
        IF bInOk AND bParaOk THEN
            fRise := fP2 - fP1;                       // 窗内压升 [帕] / Pressure rise [Pa]
            fLeakRate := fRise * fV / fWinSec;        // 压升率，分母已验正 / Rise rate, denominator verified
            IF fRise < 0.0 THEN
                bInfoBack := TRUE;                     // 反向压差（温降）信息 / Reverse rise (cooling) info
                bPass := TRUE;                         // 保守侧判合格不误杀 / Conservative pass verdict
            ELSE
                fSlack := DL_CLR_REL * MAX(ABS(fLeakLim), 1.0); // 相对余量 / Relative slack
                bPass := fLeakRate <= (fLeakLim + fSlack); // 带余量判定不做严格小于 / Slack verdict, no strict less
            END_IF
        ELSE
            fLeakRate := 0.0;                         // 异常路径确定值 / Deterministic fallback
            bPass := FALSE;                           // 异常判不合格 / Fail on invalid data
            bInfoOne := TRUE;                         // 信息级：判定拍数据非法（暂存）/ Info: illegal data at verdict, staged
        END_IF
        eState := eIdle;                              // 判定毕回待机 / Verdict done, back to idle
    eFault:
        bPass := FALSE;                               // 故障态清合格 / Fault clears verdict
        fLeakRate := 0.0;                             // 故障态清输出 / Fault clears output
        IF rTrigStart.Q AND bParaOk THEN
            eState := eStabilize;                     // 可达解除路径：重启沿重试 / Reachable release: restart edge
            uCodeLatch := 16#0000_0000;               // 清锁存码 / Clear latched code
        END_IF
    ELSE
        eState := eFault;                             // 非法状态兜底 / Illegal state fallback
        uCodeLatch := 16#0005_009B;                   // 码位：状态非法 / Code: illegal state
END_CASE

// ---- 段 5｜错误码装配：故障锁存回放优先，信息级居次 ------------------------------
IF eState = eFault THEN
    bError   := TRUE;                                 // 故障标志配对（R45）/ Fault flag paired
    uErrorId := uCodeLatch;                           // 故障码锁存回放 / Latched fault code replayed
ELSIF bInfoBack THEN
    bError   := FALSE;                                // 信息级不置故障 / Info never sets fault
    uErrorId := 16#0005_0099;                         // 信息级：反向压差判合格 / Info: reverse rise passed
ELSIF bInfoOne THEN
    bError   := FALSE;                                // 信息级不置故障 / Info never sets fault
    uErrorId := 16#0005_0099;                         // 信息级：参数/数据非法单拍回放 / Info: illegal param or data, one-scan
    bInfoOne := FALSE;                                // 发完即清 / Clear after emit
ELSE
    bError   := FALSE;                                // 无错清标志 / Clear fault flag
    uErrorId := 16#0000_0000;                         // 无码 / No code
END_IF
END_FUNCTION_BLOCK
